(* IEC 61131-3 sources: daoli-st-library/DL_Base (part 17) *)

(* ---- FB_DL_SignalQualify.st ---- *)
(*
  FB_DL_SignalQualify  —  模拟量信号有效性三态联合判定 / Analog signal qualification: over-range, frozen, wire-break
  分类 Category : DL_Base
  版本 Version  : 1.0.0
  来源 Source   : t2-1-lgf-measurement — 信号质量判定族零检索深化
  溯源 Origin   : clean-room 实现，未复制任何源码行
  功能 Function : 1) 对 fRaw 做三态联合判定：超量程（量程域外）/ 断线（低于传感器零点域）/
                  卡死（相邻拍差值持续小于卡死带超过 tFrozenTo），输出 eQual 四态枚举 + bValid；
                  2) 断线判据：fRaw < fScaleLo - fWireMargin（传感器零点域以下）→ eWireBreak；
                  3) 卡死判据：ABS(fRaw - 上拍采样) < fFrozenBand 持续 tFrozenTo → 故障级 03DC；
                  4) bReset 上升沿清全部故障锁存；判定恢复 eOk 沿置信息级码 049E。
  边界 Boundary : ① 组态闸：fScaleLo < fScaleHi 必须成立，违例置故障级 03DB，bValid 强制 FALSE；
                  ② 域判据全部使用当拍量（fRaw 与组态引脚），无锁存量自指；
                  ③ 判定派生链 IF/ELSIF/ELSE 全覆盖，枚举域防御守卫落 03DD 故障锁存；
                  ④ 无 GVL 依赖：纯引脚输入输出，无外部变量引用，无物理 IO 地址。
  依赖 Depends  : 仅 Standard.library（TON / R_TRIG）
  码表 Error codes（段 0001，窗口 03DB~03DD / 049E~04A0）:
    16#0001_03DB 故障级：量程组态非法（fScaleLo >= fScaleHi 或卡死带 <= 0），锁存至 bReset
    16#0001_03DC 故障级：信号卡死超时（冻结判据持续 tFrozenTo），锁存至 bReset
    16#0001_03DD 故障级：判定结果落枚举域外（防御守卫兜底），锁存至 bReset
    16#0001_049E 信息级：信号判定恢复正常（eQual 回 eOk 沿）
    16#0001_049F 信息级：超量程检出（伴随态）
    16#0001_04A0 信息级：断线域命中（伴随态）
  修订历史 Revision :
    2026-11-19  v1.0.0  R41 首版（批次 1 · 序号 1）
*)

TYPE E_DL_SigQual :
(
    eOk        := 0,    // 信号有效，量程域内且动态正常 / Signal valid, in range and dynamic
    eOverRange := 10,   // 超量程：超出组态量程域 / Over range, outside the configured span
    eFrozen    := 20,   // 卡死：变化量持续小于卡死带 / Frozen, change stays below the deadband
    eWireBreak := 30    // 断线：低于传感器零点域 / Wire break, below the sensor zero span
);
END_TYPE

FUNCTION_BLOCK FB_DL_SignalQualify
VAR_INPUT
    fRaw         : LREAL := 0.0;      // 原始采样值 [EU] / Raw sampled value
    fScaleLo     : LREAL := 0.0;      // 量程下限 [EU]，必须 < fScaleHi / Span lower bound
    fScaleHi     : LREAL := 100.0;    // 量程上限 [EU]，必须 > fScaleLo / Span upper bound
    fWireMargin  : LREAL := 1.0;      // 断线判据裕度 [EU]，域 >= 0 / Wire-break margin below span low
    fFrozenBand  : LREAL := 0.01;     // 卡死判定带 [EU]，域 > 0 / Frozen deadband
    tFrozenTo    : TIME := T#5S;      // 卡死确认超时 [ms]，域 > 0 / Frozen confirm timeout
    bReset       : BOOL := FALSE;     // 复位，上升沿清故障锁存 / Reset edge clears fault latches
END_VAR
VAR_OUTPUT
    eQual        : E_DL_SigQual;      // 判定结果出口 / Qualification result
    bValid       : BOOL;              // 判定有效（eOk 且无故障）/ Result usable flag
    bError       : BOOL;              // 故障锁存标志 / Fault latch flag
    nErrId       : UDINT;             // 事件码，0 = 无事件（故障锁存回放优先）/ Event code
END_VAR
VAR
    tonFrozen    : TON;               // 卡死确认定时器，无条件周期刷新 / Frozen confirm timer
    rtReset      : R_TRIG;            // 复位沿实例，无条件周期刷新 / Reset edge instance
    _fLastRaw    : LREAL := 0.0;      // 上拍采样快照 [EU] / Previous scan sample snapshot
    _fDelta      : LREAL;             // 相邻拍差值绝对值 [EU] / Absolute inter-scan delta
    _bFault      : BOOL;              // 故障锁存位（锁存量）/ Latched fault bit
    _uFault      : UDINT;             // 故障码锁存（锁存量）/ Latched fault code
    _uInfo       : UDINT;             // 信息码，每拍重算 / Transient info code
    _bOkPrev     : BOOL;              // 上拍判定有效镜像（恢复沿判据）/ Previous eOk mirror
END_VAR

(* —— 段 0：定时器与沿实例无条件周期刷新（禁置于 IF/CASE 内） —— *)
_fDelta := ABS(fRaw - _fLastRaw);                                       // 相邻拍差值（当拍量）
tonFrozen(IN := (_fDelta < fFrozenBand), PT := tFrozenTo);              // 卡死确认（每拍必调）
rtReset(CLK := bReset);                                                 // 复位沿（每拍必调）

(* —— 段 1：单拍量预清零（锁存量 _bFault/_uFault 不入清单，禁同拍抹除） —— *)
_uInfo := 16#0000_0000;             // 信息码每拍重算
bValid := FALSE;                    // 有效出口缺省 FALSE
nErrId := 16#0000_0000;             // 事件码缺省无事件
eQual := E_DL_SigQual.eOk;          // 判定缺省有效（派生链覆盖改写）

(* —— 段 2：复位沿（唯一故障解除路径，全当拍量） —— *)
IF rtReset.Q THEN                   // rtReset.Q = 当拍量
    _bFault := FALSE;               // 清故障锁存位
    _uFault := 16#0000_0000;        // 清故障锁存码
END_IF

(* —— 段 3：组态域闸（覆盖参与判据换算的全部组态引脚） —— *)
IF (fScaleLo >= fScaleHi) OR (fFrozenBand <= 0.0) OR (TIME_TO_DINT(tFrozenTo) <= 0) THEN
    _uFault := 16#0001_03DB;        // 故障级：量程组态非法
    _bFault := TRUE;
END_IF

(* —— 段 4：三态联合判定（全当拍量判据；派生链 ELSE 兜底 + 枚举域守卫） —— *)
IF NOT _bFault THEN
    IF fRaw < (fScaleLo - ABS(fWireMargin)) THEN
        eQual := E_DL_SigQual.eWireBreak;   // 断线：低于传感器零点域
        _uInfo := 16#0001_04A0;             // 信息级：断线域命中
    ELSIF (fRaw > fScaleHi) OR (fRaw < fScaleLo) THEN
        eQual := E_DL_SigQual.eOverRange;   // 超量程
        _uInfo := 16#0001_049F;             // 信息级：超量程检出
    ELSIF tonFrozen.Q THEN
        eQual := E_DL_SigQual.eFrozen;      // 卡死确认
        _uFault := 16#0001_03DC;            // 故障级：卡死超时
        _bFault := TRUE;
    ELSE
        eQual := E_DL_SigQual.eOk;          // 判定有效
        IF NOT _bOkPrev THEN
            _uInfo := 16#0001_049E;         // 信息级：判定恢复有效沿
        END_IF
    END_IF
    (* 枚举域防御守卫（等价 CASE ELSE 兜底）：判定结果必须落已知枚举域 *)
    IF (eQual <> E_DL_SigQual.eOk) AND (eQual <> E_DL_SigQual.eOverRange)
       AND (eQual <> E_DL_SigQual.eFrozen) AND (eQual <> E_DL_SigQual.eWireBreak) THEN
        _uFault := 16#0001_03DD;            // 故障级：判定态落域外
        _bFault := TRUE;
        eQual := E_DL_SigQual.eOk;          // 强制回已知态
    END_IF
END_IF

(* —— 段 5：出口单点映射（名实同源；故障锁存码回放，禁同拍抹除） —— *)
bValid := (eQual = E_DL_SigQual.eOk) AND (NOT _bFault);   // 有效出口（信息级不置故障）
IF _bFault THEN
    nErrId := _uFault;              // 故障锁存码回放
ELSE
    nErrId := _uInfo;               // 信息码
END_IF
bError := _bFault;                  // 故障标志与锁存位同源
_bOkPrev := (eQual = E_DL_SigQual.eOk);   // 恢复沿判据快照（当拍量快照）
_fLastRaw := fRaw;                  // 上拍采样快照更新（段末统一写）

END_FUNCTION_BLOCK

(* ---- FB_DL_SignalRouteMatrix.st ---- *)
//==============================================================================
// 功能块：FB_DL_SignalRouteMatrix ｜ 中文名称：2×N 可组态信号路由矩阵
// 所属子库：DL_Base ｜ 版本：v1.0.0 ｜ 日期：2026-11-23
// 兼容：CODESYS V3.5+ / TwinCAT 3 / 汇川 InoProShop（纯 IEC 61131-3，零方言）
// 功能描述：2 源 × 4 通道可组态路由矩阵：每通道独立使能 + 来源选择（源 A /
//           源 B / 空置），输出 = 使能 AND 所选源。断源哨兵：存在"通道使能
//           且已选源"但其源信号为 FALSE 时置该源断源哨兵位（正常传递同时
//           留痕，供上层诊断区分"真信号 FALSE"与"通道空置 FALSE"）。
// 开源溯源 (Origin)：原创实现（t2-1-lgf-bitlogic 位逻辑语义深化，零外部源码
//           行，clean-room 独立编写）
// 公开接口清单：输入 aSrcA / aSrcB / {bEnCh1..4, eSelCh1..4}；
//               输出 {bOutCh1..4} / bSrcALost / bSrcBLost / bValid
// 错误码表：无状态机码轨（组合路由无故障级条件）；断源诊断经
//           bSrcALost / bSrcBLost 哨兵位表达，不占用 16#0001 段码位
// 状态机：E_DL_RouteSel（本文件唯一定义，全库唯一属主）：
//           eNone = 0 / eSrcA = 1 / eSrcB = 2；非法选择值走 CASE ELSE 兜底
//           （输出 FALSE 安全侧 + 声明哨兵）
// 边界行为：① 空置通道输出恒 FALSE 且不计入断源哨兵；
//           ② 断源哨兵不屏蔽输出（传递与诊断解耦）；
//           ③ 无定时器/沿实例（纯组合逻辑，无周期刷新义务）；
//           ④ CASE 带 ELSE 非法选择值兜底（输出 FALSE 安全侧）。
// 修订历史：v1.0.0 2026-11-23 首版（R73 派单 · 批 3 · 序 13）
//==============================================================================

(*------------------------------------------------------------------------------
 * 枚举: E_DL_RouteSel（归属本功能块，同文件发布，全库唯一属主）
 * 含义: 通道来源选择，成员与 CASE 标签双向完备。
 *-----------------------------------------------------------------------------*)
TYPE E_DL_RouteSel :
(
    eNone := 0,    // 空置：通道不选源，输出恒 FALSE / Idle, no source selected
    eSrcA := 1,    // 选源 A / Source A selected
    eSrcB := 2     // 选源 B / Source B selected
);
END_TYPE

(*==============================================================================
 * 功能块: FB_DL_SignalRouteMatrix
 * 调用约定: 每个扫描周期无条件调用一次；纯组合路由，无跨拍驻留状态。
 *==============================================================================*)
FUNCTION_BLOCK FB_DL_SignalRouteMatrix
VAR_INPUT
    aSrcA   : BOOL := FALSE;           // 源 A 信号 [—] / Source A signal
    aSrcB   : BOOL := FALSE;           // 源 B 信号 [—] / Source B signal
    bEnCh1  : BOOL := FALSE;           // 通道 1 使能 / Channel 1 enable
    eSelCh1 : E_DL_RouteSel := E_DL_RouteSel.eNone; // 通道 1 来源选择 / Channel 1 source select
    bEnCh2  : BOOL := FALSE;           // 通道 2 使能 / Channel 2 enable
    eSelCh2 : E_DL_RouteSel := E_DL_RouteSel.eNone; // 通道 2 来源选择 / Channel 2 source select
    bEnCh3  : BOOL := FALSE;           // 通道 3 使能 / Channel 3 enable
    eSelCh3 : E_DL_RouteSel := E_DL_RouteSel.eNone; // 通道 3 来源选择 / Channel 3 source select
    bEnCh4  : BOOL := FALSE;           // 通道 4 使能 / Channel 4 enable
    eSelCh4 : E_DL_RouteSel := E_DL_RouteSel.eNone; // 通道 4 来源选择 / Channel 4 source select
END_VAR
VAR_OUTPUT
    bOutCh1 : BOOL;                    // 通道 1 路由输出 / Channel 1 routed output
    bOutCh2 : BOOL;                    // 通道 2 路由输出 / Channel 2 routed output
    bOutCh3 : BOOL;                    // 通道 3 路由输出 / Channel 3 routed output
    bOutCh4 : BOOL;                    // 通道 4 路由输出 / Channel 4 routed output
    bSrcALost : BOOL;                  // 断源哨兵：有通道选 A 但源 A 为 FALSE / Source-A lost sentinel
    bSrcBLost : BOOL;                  // 断源哨兵：有通道选 B 但源 B 为 FALSE / Source-B lost sentinel
    bValid  : BOOL;                    // 输出可用标志 / Outputs usable flag
END_VAR

// ---- 段 0｜出口默认值：哨兵每拍重算（组合诊断位不锁存）----
bSrcALost := FALSE;                   // 源 A 断源哨兵先清零 / Source-A lost sentinel cleared first
bSrcBLost := FALSE;                   // 源 B 断源哨兵先清零 / Source-B lost sentinel cleared first
bValid    := TRUE;                    // 可用标志默认 TRUE / Usable flag preset TRUE

// ---- 段 1｜通道 1/2 路由（CASE 带 ELSE；空置与非法值安全侧输出 FALSE）----
CASE eSelCh1 OF                       // 通道 1 来源判决 / Channel 1 source decision
    E_DL_RouteSel.eNone:               // 空置：输出 FALSE，不计哨兵 / Idle, FALSE, no sentinel
        bOutCh1 := FALSE;              // 通道 1 输出 / Channel 1 output
    E_DL_RouteSel.eSrcA:               // 选源 A：使能闸 + 断源哨兵留痕 / Source A, enable gate plus lost sentinel
        bOutCh1 := bEnCh1 AND aSrcA;   // 通道 1 输出 / Channel 1 output
        bSrcALost := bSrcALost OR (bEnCh1 AND NOT aSrcA); // 断源哨兵累积 / Lost sentinel accumulate
    E_DL_RouteSel.eSrcB:               // 选源 B：使能闸 + 断源哨兵留痕 / Source B, enable gate plus lost sentinel
        bOutCh1 := bEnCh1 AND aSrcB;   // 通道 1 输出 / Channel 1 output
        bSrcBLost := bSrcBLost OR (bEnCh1 AND NOT aSrcB); // 断源哨兵累积 / Lost sentinel accumulate
    ELSE                               // 非法选择值兜底（R21：CASE 必带 ELSE）
        bOutCh1 := FALSE;              // 安全侧输出 FALSE / Safe-side FALSE output
END_CASE
CASE eSelCh2 OF                       // 通道 2 来源判决 / Channel 2 source decision
    E_DL_RouteSel.eNone:               // 空置：输出 FALSE，不计哨兵 / Idle, FALSE, no sentinel
        bOutCh2 := FALSE;              // 通道 2 输出 / Channel 2 output
    E_DL_RouteSel.eSrcA:               // 选源 A：使能闸 + 断源哨兵留痕 / Source A, enable gate plus lost sentinel
        bOutCh2 := bEnCh2 AND aSrcA;   // 通道 2 输出 / Channel 2 output
        bSrcALost := bSrcALost OR (bEnCh2 AND NOT aSrcA); // 断源哨兵累积 / Lost sentinel accumulate
    E_DL_RouteSel.eSrcB:               // 选源 B：使能闸 + 断源哨兵留痕 / Source B, enable gate plus lost sentinel
        bOutCh2 := bEnCh2 AND aSrcB;   // 通道 2 输出 / Channel 2 output
        bSrcBLost := bSrcBLost OR (bEnCh2 AND NOT aSrcB); // 断源哨兵累积 / Lost sentinel accumulate
    ELSE                               // 非法选择值兜底（R21：CASE 必带 ELSE）
        bOutCh2 := FALSE;              // 安全侧输出 FALSE / Safe-side FALSE output
END_CASE

// ---- 段 2｜通道 3/4 路由（同段 1 口径）----
CASE eSelCh3 OF                       // 通道 3 来源判决 / Channel 3 source decision
    E_DL_RouteSel.eNone:               // 空置：输出 FALSE，不计哨兵 / Idle, FALSE, no sentinel
        bOutCh3 := FALSE;              // 通道 3 输出 / Channel 3 output
    E_DL_RouteSel.eSrcA:               // 选源 A：使能闸 + 断源哨兵留痕 / Source A, enable gate plus lost sentinel
        bOutCh3 := bEnCh3 AND aSrcA;   // 通道 3 输出 / Channel 3 output
        bSrcALost := bSrcALost OR (bEnCh3 AND NOT aSrcA); // 断源哨兵累积 / Lost sentinel accumulate
    E_DL_RouteSel.eSrcB:               // 选源 B：使能闸 + 断源哨兵留痕 / Source B, enable gate plus lost sentinel
        bOutCh3 := bEnCh3 AND aSrcB;   // 通道 3 输出 / Channel 3 output
        bSrcBLost := bSrcBLost OR (bEnCh3 AND NOT aSrcB); // 断源哨兵累积 / Lost sentinel accumulate
    ELSE                               // 非法选择值兜底（R21：CASE 必带 ELSE）
        bOutCh3 := FALSE;              // 安全侧输出 FALSE / Safe-side FALSE output
END_CASE
CASE eSelCh4 OF                       // 通道 4 来源判决 / Channel 4 source decision
    E_DL_RouteSel.eNone:               // 空置：输出 FALSE，不计哨兵 / Idle, FALSE, no sentinel
        bOutCh4 := FALSE;              // 通道 4 输出 / Channel 4 output
    E_DL_RouteSel.eSrcA:               // 选源 A：使能闸 + 断源哨兵留痕 / Source A, enable gate plus lost sentinel
        bOutCh4 := bEnCh4 AND aSrcA;   // 通道 4 输出 / Channel 4 output
        bSrcALost := bSrcALost OR (bEnCh4 AND NOT aSrcA); // 断源哨兵累积 / Lost sentinel accumulate
    E_DL_RouteSel.eSrcB:               // 选源 B：使能闸 + 断源哨兵留痕 / Source B, enable gate plus lost sentinel
        bOutCh4 := bEnCh4 AND aSrcB;   // 通道 4 输出 / Channel 4 output
        bSrcBLost := bSrcBLost OR (bEnCh4 AND NOT aSrcB); // 断源哨兵累积 / Lost sentinel accumulate
    ELSE                               // 非法选择值兜底（R21：CASE 必带 ELSE）
        bOutCh4 := FALSE;              // 安全侧输出 FALSE / Safe-side FALSE output
END_CASE

// ---- 段 3｜统一出口：可用标志（纯组合无防御失败路径）----
bValid := TRUE;                       // 组合路由恒可用 / Combinational routing always usable
END_FUNCTION_BLOCK

(* ---- FB_DL_SignalSeqGuard.st ---- *)
(*
  ==================================================================
  组件名 Component  : FB_DL_SignalSeqGuard
  分类   Category   : DL_Base
  复杂度 Complexity  : cx3
  版本   Version    : 1.0.0
  功能   Purpose    : 多路信号到达顺序守卫。N = 4 路布尔信号按期望序（ENUM 四选一：
                      升序 1→2→3→4 / 降序 4→3→2→1 / 对 1→2 / 对 3→4）在 tWindow
                      内逐沿校验到达顺序；乱序即置 eFault = eOrderViolation 并锁存，
                      窗内未完成置 eWindowTimeout；正常序完成置 bSeqOk 单拍脉冲。
                      复位上升沿清全部锁存。同拍多沿按 1..4 固定序检查（确定性口径）。
  来源   Source     : t2-1-lgf-converter
  溯源   Origin     : IEC 61131-3 标准语义的道莅防御性实现；到达顺序校验为通用
                      联锁语义，clean-room 自研实现，未复制任何闭源代码行。
  平台   Platform   : 纯 IEC 61131-3（TON / R_TRIG / ARRAY，无私有库）
  作者   Author     : 道莅代码库 · PLC 编程专家（R56）
  ------------------------------------------------------------------
  边界 Boundary     :
                      一 本件只做到达顺序校验，不产生任何输出命令（属主边界）；
                      二 eWait 类相（eRun）退出条件 ≥2 条：完成沿 / 超时 / 乱序 /
                         失能，四条并列（R98）；
                      三 序列表在组态相一次性落定，乱序判据只用序表与步进游标；
                      四 故障锁存解除路径 = bReset 上升沿（唯一路径，头注释声明，R188）；
                      五 无全局变量、无外部变量声明、无物理地址寻址。
  输出契约 Output contract:
                      bSeqOk 为单拍脉冲（内部 _bOkInt 置位、统一出口映射后撤销，R187）；
                      eFault 为锁存回放；eModeBad 为模式枚举非法兜底（R128）。
  修订记录 Revision  :
    2026-11-20  v1.0.0  R56 首版（批 2 · 序号 7）
  ==================================================================
*)

TYPE E_DL_SsgMode :
(
    eAscending  := 0, // 升序：1→2→3→4 / ascending, one to four
    eDescending := 1, // 降序：4→3→2→1 / descending, four to one
    ePair12     := 2, // 对序：1→2 / pair order, one then two
    ePair34     := 3  // 对序：3→4 / pair order, three then four
);
END_TYPE

TYPE E_DL_SsgPhase :
(
    eIdle  := 0,  // 空闲：等待启动 / idle, waiting for the start
    eRun   := 10, // 校验中：逐沿核对到达顺序 / running, the arrivals are checked edge by edge
    eDone  := 20, // 完成：顺序通过，驻留一拍 / done, the order passed and the phase holds one scan
    eFault := 90  // 故障：成因锁存 / fault, the cause is latched
);
END_TYPE

TYPE E_DL_SsgFault :
(
    eNone          := 0, // 无成因 / no cause
    eOrderViolation:= 1, // 到达顺序违例（故障级，与 bError 配对）/ the arrival order was violated, fault grade paired with bError
    eWindowTimeout := 2, // 时窗内未完成（故障级，与 bError 配对）/ the window expired without completion, fault grade paired with bError
    eModeBad       := 3, // 模式枚举非法（故障级，与 bError 配对）/ the mode enumeration is illegal, fault grade paired with bError
    ePhaseBad      := 4  // 非法相位兜底（故障级，与 bError 配对）/ illegal phase fallback, fault grade paired with bError
);
END_TYPE

FUNCTION_BLOCK FB_DL_SignalSeqGuard
VAR_INPUT
    bEnable   : BOOL := TRUE;    // 使能，失能时停校验回空闲 [-] / enable, the check stops when disabled
    bReset    : BOOL := FALSE;   // 复位上升沿清全部锁存 [-] / reset rising edge clears every latch
    bIn1      : BOOL := FALSE;   // 信号 1 [-] / signal one
    bIn2      : BOOL := FALSE;   // 信号 2 [-] / signal two
    bIn3      : BOOL := FALSE;   // 信号 3 [-] / signal three
    bIn4      : BOOL := FALSE;   // 信号 4 [-] / signal four
    eSeqMode  : E_DL_SsgMode := E_DL_SsgMode.eAscending; // 期望到达序 [枚举] / the expected arrival order [enum]
    tWindow   : TIME := T#2S;    // 到达顺序时窗 [毫秒]，域 大于零 / arrival order window [millisecond], domain above zero
END_VAR
VAR_OUTPUT
    bSeqOk    : BOOL := FALSE; // 顺序通过单拍脉冲 [-] / the order passed single shot pulse
    nStep     : INT := 0;      // 已到位步数 [步] / the arrived step count [step]
    ePhase    : E_DL_SsgPhase := E_DL_SsgPhase.eIdle; // 相位出口 [枚举] / phase outlet [enum]
    eFault    : E_DL_SsgFault := E_DL_SsgFault.eNone; // 成因出口，锁存回放 [枚举] / cause outlet replayed from the latch [enum]
    bError    : BOOL := FALSE; // 故障锁存标志 [-] / fault latch flag
END_VAR
VAR
    rtIn1     : R_TRIG;  // 信号 1 沿检测，段 0 无条件刷新 / signal one edge, refreshed unconditionally in segment zero
    rtIn2     : R_TRIG;  // 信号 2 沿检测，段 0 无条件刷新 / signal two edge, refreshed unconditionally in segment zero
    rtIn3     : R_TRIG;  // 信号 3 沿检测，段 0 无条件刷新 / signal three edge, refreshed unconditionally in segment zero
    rtIn4     : R_TRIG;  // 信号 4 沿检测，段 0 无条件刷新 / signal four edge, refreshed unconditionally in segment zero
    rtReset   : R_TRIG;  // 复位沿检测，段 0 无条件刷新 / reset edge, refreshed unconditionally in segment zero
    tonWindow : TON;     // 到达顺序时窗，段 0 无条件刷新 / arrival window timer, refreshed unconditionally in segment zero
    _ePhase   : E_DL_SsgPhase := E_DL_SsgPhase.eIdle; // 内部相位，CASE 唯一写入目标 / internal phase, the only CASE write target
    _eFaulC   : E_DL_SsgFault := E_DL_SsgFault.eNone; // 故障级成因，锁存至复位沿 / fault cause, latched until the reset edge
    _bFault   : BOOL := FALSE; // 故障锁存位 [-] / fault latch bit
    _bInit    : BOOL := FALSE; // 首扫初始化完成标志（R310）/ first scan initialisation flag
    _bOkInt   : BOOL := FALSE; // 通过脉冲内部位，统一出口映射 / internal passed bit, mapped at the unified outlet
    _nStep    : INT := 0;      // 已到位步数 [步] / the arrived step count [step]
    _nSeqLen  : INT := 4;      // 序列长度（四序或两序）[步] / the sequence length, four or two steps
    _nSig     : INT := 0;      // 本拍到沿的信号号 [信号号] / the signal number that edged this scan
    _anOrder  : ARRAY[1..4] OF INT := [0, 0, 0, 0]; // 期望到达序表（0 = 空槽）[信号号] / the expected order table, zero is an empty slot
END_VAR

// 段 0｜定时器与沿检测无条件周期刷新（禁入分支），IN 只串相位闸与故障闸（FB50-1）/ segment 0, unconditional refresh, no instance call inside a branch
rtIn1(CLK := bIn1); // 信号 1 沿 / the signal one edge
rtIn2(CLK := bIn2); // 信号 2 沿 / the signal two edge
rtIn3(CLK := bIn3); // 信号 3 沿 / the signal three edge
rtIn4(CLK := bIn4); // 信号 4 沿 / the signal four edge
rtReset(CLK := bReset); // 复位沿 / the reset edge
tonWindow(IN := (_ePhase = E_DL_SsgPhase.eRun) AND (NOT _bFault), PT := tWindow); // 到达顺序时窗，IN 串校验相闸与故障闸 / the arrival window with the phase and fault gates on IN

// 段 1｜首扫初始化（R310）/ segment 1, first scan initialisation
IF NOT _bInit THEN // 首扫一拍 / the very first scan
    _bInit := TRUE; // 置首扫完成标志 / raise the first scan flag
    _ePhase := E_DL_SsgPhase.eIdle; // 相位从空闲起步 / the phase starts from idle
    _eFaulC := E_DL_SsgFault.eNone; // 故障级成因清零 / clear the fault cause
    _bFault := FALSE; // 故障锁存清零 / clear the fault latch
    _nStep := 0; // 步数清零 / clear the step count
END_IF

// 段 2｜复位沿作用域：清锁存 / 迁相位 / 清步数（三项逐项声明）/ segment 2, reset edge scope declared item by item
IF rtReset.Q THEN // 复位沿 / the reset edge
    _bFault := FALSE; // 作用域一：清故障锁存 / scope one, clear the fault latch
    _eFaulC := E_DL_SsgFault.eNone; // 作用域一：清故障级成因 / scope one, clear the fault cause
    _ePhase := E_DL_SsgPhase.eIdle; // 作用域二：迁回空闲相 / scope two, migrate back to idle
    _nStep := 0; // 作用域三：清步数 / scope three, clear the step count
END_IF

// 段 3｜序表组态：按模式一次性落定，非法模式判故障 / segment 3, the order table settles per the mode, an illegal mode faults
CASE eSeqMode OF // 模式分派 / the mode dispatch
E_DL_SsgMode.eAscending: // 升序 / ascending
    _anOrder[1] := 1; // 第一位信号 1 / the first slot takes signal one
    _anOrder[2] := 2; // 第二位信号 2 / the second slot takes signal two
    _anOrder[3] := 3; // 第三位信号 3 / the third slot takes signal three
    _anOrder[4] := 4; // 第四位信号 4 / the fourth slot takes signal four
    _nSeqLen := 4; // 序列长度四 / the length is four
E_DL_SsgMode.eDescending: // 降序 / descending
    _anOrder[1] := 4; // 第一位信号 4 / the first slot takes signal four
    _anOrder[2] := 3; // 第二位信号 3 / the second slot takes signal three
    _anOrder[3] := 2; // 第三位信号 2 / the third slot takes signal two
    _anOrder[4] := 1; // 第四位信号 1 / the fourth slot takes signal one
    _nSeqLen := 4; // 序列长度四 / the length is four
E_DL_SsgMode.ePair12: // 对序 1→2 / pair one then two
    _anOrder[1] := 1; // 第一位信号 1 / the first slot takes signal one
    _anOrder[2] := 2; // 第二位信号 2 / the second slot takes signal two
    _anOrder[3] := 0; // 空槽 / an empty slot
    _anOrder[4] := 0; // 空槽 / an empty slot
    _nSeqLen := 2; // 序列长度二 / the length is two
E_DL_SsgMode.ePair34: // 对序 3→4 / pair three then four
    _anOrder[1] := 3; // 第一位信号 3 / the first slot takes signal three
    _anOrder[2] := 4; // 第二位信号 4 / the second slot takes signal four
    _anOrder[3] := 0; // 空槽 / an empty slot
    _anOrder[4] := 0; // 空槽 / an empty slot
    _nSeqLen := 2; // 序列长度二 / the length is two
ELSE // 非法模式兜底（R128）/ the illegal mode fallback
    IF (NOT _bFault) AND (_ePhase <> E_DL_SsgPhase.eFault) THEN // 未锁存才迁移（防同拍抹除）/ migrate only while unlatched
        _bFault := TRUE; // 置故障锁存 / raise the fault latch
        _eFaulC := E_DL_SsgFault.eModeBad; // 故障级成因（R45 配对 bError）/ the fault cause paired with bError
        _ePhase := E_DL_SsgPhase.eFault; // 迁故障相 / migrate to the fault phase
    END_IF
END_CASE

// 段 4｜本拍到沿信号号判定：同拍多沿按 1..4 固定序（确定性口径）/ segment 4, the edged signal number, multiple edges resolve in the fixed one to four order
_nSig := 0; // 信号号预置零 / preset the signal number to zero
IF rtIn1.Q THEN // 信号 1 到沿 / signal one edged
    _nSig := 1; // 记信号 1 / take signal one
ELSIF rtIn2.Q THEN // 信号 2 到沿 / signal two edged
    _nSig := 2; // 记信号 2 / take signal two
ELSIF rtIn3.Q THEN // 信号 3 到沿 / signal three edged
    _nSig := 3; // 记信号 3 / take signal three
ELSIF rtIn4.Q THEN // 信号 4 到沿 / signal four edged
    _nSig := 4; // 记信号 4 / take signal four
END_IF

// 段 5｜相位机：ENUM + CASE，含 ELSE 非法相位兜底（R128）/ segment 5, the phase machine with an ELSE fallback
CASE _ePhase OF
E_DL_SsgPhase.eIdle: // 空闲相：使能且无故障即起校验 / idle, the check starts when enabled and unfaulted
    IF bEnable AND (NOT _bFault) THEN // 使能且无故障 / enabled and unfaulted
        _nStep := 0; // 步数清零 / clear the step count
        _ePhase := E_DL_SsgPhase.eRun; // 迁校验相 / migrate to the run phase
    END_IF

E_DL_SsgPhase.eRun: // 校验相：逐沿核对到达顺序（退出条件 ≥2：完成 / 超时 / 乱序 / 失能，R98）/ the run phase with at least two exit conditions
    nStep := _nStep; // 步数出口跟随 / the step outlet follows
    IF NOT bEnable THEN // 失能 / disabled
        _ePhase := E_DL_SsgPhase.eIdle; // 回空闲相 / return to idle
    ELSIF tonWindow.Q THEN // 时窗耗尽未完成 / the window expired without completion
        _bFault := TRUE; // 置故障锁存 / raise the fault latch
        _eFaulC := E_DL_SsgFault.eWindowTimeout; // 故障级成因（R45 配对 bError）/ the fault cause paired with bError
        _ePhase := E_DL_SsgPhase.eFault; // 迁故障相 / migrate to the fault phase
    ELSIF _nSig > 0 THEN // 本拍有信号到沿 / a signal edged this scan
        IF _nSig = _anOrder[_nStep + 1] THEN // 与期望序位一致 / the arrival matches the expected slot
            _nStep := _nStep + 1; // 步数推进 / advance the step
            IF _nStep >= _nSeqLen THEN // 序列完成 / the sequence is complete
                _bOkInt := TRUE; // 通过脉冲内部位置位（统一出口映射，R187）/ raise the internal passed bit, mapped at the unified outlet
                _ePhase := E_DL_SsgPhase.eDone; // 迁完成相 / migrate to the done phase
            END_IF
        ELSE // 乱序 / an out of order arrival
            _bFault := TRUE; // 置故障锁存 / raise the fault latch
            _eFaulC := E_DL_SsgFault.eOrderViolation; // 故障级成因（R45 配对 bError）/ the fault cause paired with bError
            _ePhase := E_DL_SsgPhase.eFault; // 迁故障相 / migrate to the fault phase
        END_IF
    END_IF

E_DL_SsgPhase.eDone: // 完成相：脉冲已交付（拍 N 进入：序到位 / 本拍行为：脉冲映射 / 拍 N+1 转出：无条件回空闲，R80 三段）/ the done phase, the pulse was delivered
    _ePhase := E_DL_SsgPhase.eIdle; // 无条件回空闲相准备下一轮（失能态下同样回到空闲语义）/ back to idle for the next round unconditionally, the same idle semantics under a disable

E_DL_SsgPhase.eFault: // 故障相：成因锁存，等待复位沿 / the fault phase, the cause is latched until the reset edge
    nStep := _nStep; // 步数出口冻结保持 / the step outlet holds frozen

ELSE // 非法相位兜底（R128）/ the illegal phase fallback
    _bFault := TRUE; // 置故障锁存 / raise the fault latch
    _eFaulC := E_DL_SsgFault.ePhaseBad; // 故障级成因（R45 配对 bError）/ the fault cause paired with bError
    _ePhase := E_DL_SsgPhase.eFault; // 迁故障相 / migrate to the fault phase
END_CASE

// 段 6｜统一出口 / segment 6, the unified outlet
bSeqOk := _bOkInt; // 通过脉冲映射本拍值 / map the passed pulse for this scan
_bOkInt := FALSE; // 映射后立即撤销，保证单拍宽度（R187 两段式）/ revoke right after mapping to keep a single scan width
nStep := _nStep; // 步数出口 / the step outlet
ePhase := _ePhase; // 相位出口单点映射 / single point phase outlet mapping
eFault := _eFaulC; // 成因出口锁存回放 / the cause outlet replayed from the latch
bError := _bFault; // 故障标志与锁存位同源 / the fault flag shares the latch source
END_FUNCTION_BLOCK

(* ---- FB_DL_SignalStagnationWatch.st ---- *)
(*
  ==================================================================
  组件名 Component  : FB_DL_SignalStagnationWatch
  分类   Category   : DL_Base
  复杂度 Complexity  : cx3
  版本   Version    : 1.0.0
  功能   Purpose    : 信号呆滞（卡死）检测。双判据持续 tStall 判呆滞：
                      ① 值纹波消失——相邻拍变化量 |Δ| ≤ fEps 持续；
                      ② 伴生活动信号边沿计数归零——活动观测窗内零边沿。
                      两判据同时成立才出呆滞电平与单拍事件。
  来源   Source     : iec-std-wrapper（T0）
  溯源   Origin     : IEC 61131-3 标准语义的道莅防御性实现；呆滞双判据为公开
                      诊断语义，clean-room 自研实现，未复制任何闭源代码行。
  平台   Platform   : 纯 IEC 61131-3（Standard.library: TON / R_TRIG，无私有库）
  分工声明 Split     : 与 FB_DL_SignalDebounce 分工——Debounce 是（抑制）件
                      （吸收毛刺防误动），本件是（检出）件（发现信号呆滞
                      疑点），方向相反、互不替代；与 FB_DL_SensorDropoutHold
                      分工——掉线保持件处理无效值，本件处理有效但不动值。
  作者   Author     : 道莅代码库 · PLC 编程专家（R57）
  ------------------------------------------------------------------
  边界 Boundary     :
                      一 fEps 为显式纹波死区参数，组态闸要求 > 0（信息级）；
                      二 tStall 期间边沿计数窗独立自复位（R188：IN := NOT Q），
                         与呆滞计时互不牵连；
                      三 使能断开即复位：计时清零、窗计数清零、出口回假，
                         不锁存（每拍重算）；
                      四 首扫快照取当拍，无假呆滞（tonStall 从零起步）；
                      五 无全局变量、无外部变量声明、无物理地址寻址。
  修订记录 Revision  :
    2026-11-21  v1.0.0  R57 首版（批 1 · 序号 4）
  ==================================================================
*)

FUNCTION_BLOCK FB_DL_SignalStagnationWatch
VAR_INPUT
    fValue    : LREAL := 0.0;    // 被监视值 [工程单位] / the monitored value [engineering unit]
    bActivity : BOOL := FALSE;   // 伴生活动信号（如传感器自检翻转）[-] / the companion activity signal
    fEps      : LREAL := 0.01;   // 纹波死区 [工程单位]，域 大于零 / the ripple deadband [engineering unit], above zero
    tStall    : TIME := T#10S;   // 呆滞确认窗 [毫秒] / the stall confirm window [millisecond]
    tEdgeWin  : TIME := T#5S;    // 边沿观测窗 [毫秒] / the edge observation window [millisecond]
    bEnable   : BOOL := TRUE;    // 使能，失能即复位不锁存 [-] / enable, disabling resets without latching
    bReset    : BOOL := FALSE;   // 复位上升沿清计数 [-] / reset rising edge clears the counters
END_VAR
VAR_OUTPUT
    bStalled    : BOOL := FALSE; // 呆滞电平出口（双判据同时成立）[-] / the stalled level outlet, both criteria met
    bStallEvent : BOOL := FALSE; // 呆滞进入单拍事件 [-] / the stall entry one-scan event
    nRippleCnt  : UDINT := 0;    // 纹波事件累计 [次] / the ripple event count [count]
    nActWinCnt  : UDINT := 0;    // 当前观测窗内活动边沿计数 [次] / the activity edge count in the current window [count]
    uErrorId    : UDINT := 0;    // 信息级码，0 = 正常 / informational code, zero is ok
    bError      : BOOL := FALSE; // 信息级错误标志（每拍重算）/ informational flag, recomputed each scan
END_VAR
VAR
    rtReset : R_TRIG;  // 复位沿检测，段 0 无条件刷新 / the reset edge, refreshed unconditionally
    rtAct   : R_TRIG;  // 活动信号沿检测，段 0 无条件刷新 / the activity edge, refreshed unconditionally
    rtStall : R_TRIG;  // 呆滞电平沿检测，段 0 无条件刷新 / the stalled level edge, refreshed unconditionally
    tonStall: TON;     // 呆滞确认窗，段 0 无条件刷新 / the stall confirm timer, refreshed unconditionally
    tonWin  : TON;     // 边沿观测窗（自复位），段 0 无条件刷新 / the observation window, self resetting, refreshed unconditionally
    _bInit  : BOOL := FALSE; // 首扫初始化完成标志（R310）/ first scan flag
    _fPrev  : LREAL := 0.0;  // 上拍值快照 [工程单位] / previous scan value snapshot [engineering unit]
    _bRipple: BOOL := FALSE; // 本拍纹波事件标记（上拍值供段 0 判据闸使用）/ the ripple flag this scan, the last value feeds the segment zero gate
    _bCfgOk : BOOL := FALSE; // 组态域内 [-] / the configuration inside the domain
END_VAR

// 段 0｜定时器与沿检测无条件周期刷新（禁入分支）；观测窗自复位（R188）/ segment 0, unconditional refresh, the window self resetting
rtReset(CLK := bReset); // 复位沿 / the reset edge
rtAct(CLK := bActivity); // 活动沿 / the activity edge
rtStall(CLK := bStalled); // 呆滞电平沿 / the stalled level edge
tonStall(IN := _bCfgOk AND bEnable AND (NOT _bRipple) AND (rtAct.Q = FALSE) AND (nActWinCnt = 0), PT := tStall); // 呆滞窗，IN 串双判据闸 / the stall timer gated by both criteria
tonWin(IN := bEnable AND (NOT tonWin.Q), PT := tEdgeWin); // 观测窗自复位循环（R188）/ the self resetting observation loop

// 段 1｜首扫初始化（R310）：快照取当拍防假呆滞 / segment 1, first scan, the snapshot takes this scan
IF NOT _bInit THEN // 首扫一拍 / the first scan
    _bInit := TRUE; // 置首扫标志 / raise the flag
    _fPrev := fValue; // 快照取当拍 / the snapshot takes this scan
END_IF

// 段 2｜复位沿作用域：清计数（出口电平随计时自清，无需另清）/ segment 2, reset edge scope
IF rtReset.Q THEN // 复位沿 / the reset edge
    nRippleCnt := 0; // 清纹波计数 / clear the ripple counter
    nActWinCnt := 0; // 清窗计数 / clear the window counter
END_IF

// 段 3｜组态域闸（信息级，每拍重算）/ segment 3, the configuration gate, informational
_bCfgOk := (fEps > 0.0) AND (fEps = fEps) AND ((fEps - fEps) = (fEps - fEps)) AND (tStall > T#0S) AND (tEdgeWin > T#0S); // 死区与窗域判定 / the deadband and window verdict
IF NOT _bCfgOk THEN // 组态非法 / an illegal configuration
    uErrorId := 16#0001_0001; // 信息级：组态越域 / informational, a config violation
    bError   := TRUE; // 置信息级标志 / raise the flag
ELSE // 域内 / inside the domain
    uErrorId := 16#0000_0000; // 正常码 / the ok code
    bError   := FALSE; // 清标志 / clear the flag
END_IF

// 段 4｜双判据量测 / segment 4, the dual criteria measurement
_bRipple := ABS(fValue - _fPrev) > fEps; // 纹波判据（变化量超死区）/ the ripple verdict beyond the deadband
IF _bRipple THEN // 纹波事件 / a ripple event
    nRippleCnt := nRippleCnt + 1; // 纹波计数推进 / advance the ripple counter
    IF nRippleCnt = 4294967295 THEN // UDINT 上界防回绕 / the wrap guard
        nRippleCnt := 4294967294; // 钳在次上界 / clamp below the ceiling
    END_IF
END_IF
IF rtAct.Q THEN // 活动沿 / an activity edge
    nActWinCnt := nActWinCnt + 1; // 窗内计数推进 / advance the window counter
END_IF
IF tonWin.Q THEN // 观测窗到期：窗计数独立归零重开（边界二）/ the window expired, the counter reset independently
    nActWinCnt := 0; // 窗计数归零 / the window counter zeroed
END_IF
IF NOT bEnable THEN // 失能即复位不锁存（边界三）/ disabled resets without latching
    nRippleCnt := 0; // 清纹波计数 / clear the ripple counter
    nActWinCnt := 0; // 清窗计数 / clear the window counter
END_IF

// 段 5｜统一出口：双判据电平 + 进入事件 / segment 5, the unified outlet
bStalled := _bCfgOk AND bEnable AND tonStall.Q AND (nActWinCnt = 0); // 双判据电平 / the dual criteria level
bStallEvent := rtStall.Q; // 进入单拍事件（沿检测已无条件刷新）/ the entry one-scan event
IF NOT bEnable THEN // 失能拍出口回假 / the disabled scan forces false
    bStalled := FALSE; // 电平回假 / the level false
    bStallEvent := FALSE; // 事件回假 / the event false
END_IF
_fPrev := fValue; // 快照推进（无条件）/ the snapshot advances unconditionally
END_FUNCTION_BLOCK

(* ---- FB_DL_SignalStuckWatch.st ---- *)
(*
  Name        : FB_DL_SignalStuckWatch
  Category    : DL_Base
  Version     : 1.0.0
  Purpose     : 信号卡死监视：监视值在卡死判定窗内变化量始终不超过死区（变化率恒零）即报警，捕捉传感器冻结/线束搭死；/ Signal stuck watch: raises an alarm when the monitored value stays within the deadband for the whole stuck window, catching frozen sensors or shorted wiring
  溯源        : 借 t2-1-lgf 的分类/参数域组织，clean-room 实现
  Boundary    : ① 组态闸：死区 < 0 / 卡死窗 <= T#0S → 锁存故障（死区 0 合法：严格等值判死）；
                ② 卡死判定窗用 TON，IN 由「未变化 + 已取基线」派生并串 eMon 相位闸（族③：eIdle/eFault 不计时，上拍相位 1 拍延迟可接受），段 0 无 IF 包裹；
                ③ 非有限值该拍不更新基线不计时（防 NaN 把窗持续清零而漏报，也防污染基线）；
                ④ 基线快照在迁入 eMon 拍取（fValue 首值），变化超死区即刷新基线并重置计时；
                ⑤ bStuck 锁存至复位沿；bStuck 起始沿单拍脉冲 bStuckEdge 供事件记录（R187 两段式）。
*)
TYPE E_DL_SswState :
(
    eIdle  := 0,                             (* 未使能 / Disabled *)
    eMon   := 10,                            (* 卡死监视运行 / Monitoring *)
    eFault := 90                             (* 故障锁存相 / Fault latched *)
);
END_TYPE

TYPE E_DL_SswCause :
(
    eNone       := 0,                        (* 无故障成因 / No cause *)
    eCfgIllegal := 1,                        (* 组态非法：死区/窗口越域 / Illegal config *)
    eStuck      := 2,                        (* 信号卡死（窗满无有效变化） / Signal stuck *)
    ePhaseBad   := 3                         (* 非法相位兜底 / Illegal phase fallback *)
);
END_TYPE

FUNCTION_BLOCK FB_DL_SignalStuckWatch
VAR_INPUT
    fValue    : REAL := 0.0;                 (* 被监视信号值（任意工程量）[-] / Monitored signal value *)
    fDeadband : REAL := 0.01;               (* 变化判定死区，域 >= 0 [工程单位] / Deadband for change detection *)
    tStuckWin : TIME := T#60S;              (* 卡死判定窗长，域 > T#0S [ms] / Stuck window length, > 0 *)
    bEnable   : BOOL := TRUE;               (* 监视使能 [-] / Enable *)
    bReset    : BOOL := FALSE;              (* 复位命令，上升沿清报警与故障 [-] / Reset command *)
END_VAR
VAR_OUTPUT
    fDelta    : REAL;                        (* 本拍相对基线变化量（实时派生）[工程单位] / Delta versus baseline *)
    bStuck    : BOOL;                        (* 卡死报警锁存（复位沿清）[-] / Stuck alarm latched *)
    bStuckEdge: BOOL;                        (* 卡死报警起始沿（单拍脉冲）[-] / Stuck alarm rising edge pulse *)
    fLastMove : TIME;                       (* 最近一次有效变化距今时长（本窗计时镜像）[ms] / Time since last valid move *)
    eState    : E_DL_SswState;               (* 状态出口 / State outlet *)
    eCause    : E_DL_SswCause;               (* 故障成因出口（R190 归因唯一） / Fault cause outlet *)
    bError    : BOOL;                        (* 故障锁存标志 [-] / Fault latch flag *)
END_VAR
VAR
    _eState   : E_DL_SswState := E_DL_SswState.eIdle;    (* 内部相位（CASE 唯一写入目标） / Internal phase *)
    _eCause   : E_DL_SswCause := E_DL_SswCause.eNone;    (* 故障成因锁存量 / Latched cause *)
    rtReset   : R_TRIG;                      (* 复位沿实例，段 0 无条件调用 / Reset edge instance *)
    rtStuck   : R_TRIG;                      (* 卡死计时器输出沿实例，段 0 无条件调用 / Stuck-timer edge instance *)
    tonStuck  : TON;                         (* 卡死判定窗计时器（IN 由变化判据派生 + 相位闸） / Stuck window timer *)
    _bFault   : BOOL;                        (* 故障锁存位 / Latched fault bit *)
    _bCfgBad  : BOOL;                        (* 组态非法当拍量 / Illegal config this scan *)
    _bFin     : BOOL;                        (* 监视值有限性当拍量 / Value finiteness *)
    _bMoved   : BOOL;                        (* 本拍有效变化当拍量（超死区） / Valid move this scan *)
    _bSeen    : BOOL;                        (* 基线已建立标志 / Baseline established flag *)
    _fLast    : REAL;                        (* 基线快照（最近一次有效变化的值）[工程单位] / Baseline snapshot *)
    _fDeltaI  : REAL;                        (* 变化量中间量 [工程单位] / Delta intermediate *)
    _bStuckC  : BOOL;                        (* 卡死起始沿内部单拍量（出口统一映射，R187） / Stuck-edge internal pulse *)
END_VAR
VAR CONSTANT
    DL_SSW_EPS : REAL := 1.0E-6;             (* 判零容差（REAL 量级）[-] / Epsilon *)
END_VAR

(* —— 段 0：当拍判据派生 + 实例无条件刷新（R228A；R_TRIG/TON 全在段 0，无 IF 包裹） —— *)
_bCfgBad := (fDeadband < 0.0) OR NOT (tStuckWin > T#0S);                       (* 死区非负闸 + 卡死窗正域闸 / Deadband and window gates *)
rtReset(CLK := bReset);                                                        (* 复位沿每拍必调 / Reset edge every scan *)
_bFin := (fValue = fValue) AND ((fValue - fValue) = (fValue - fValue));        (* 监视值 NaN 自反 + Inf 差判闸 / Value NaN and Inf gate *)
_fDeltaI := fValue - _fLast;                                                   (* 相对基线变化量（基线无效期不用于判据）[工程单位] / Delta versus baseline *)
_bMoved := _bFin AND _bSeen AND (ABS(_fDeltaI) > fDeadband);                   (* 有效变化：有限 + 基线在 + 超死区（死区 0 即严格不等） / Valid move gate *)
tonStuck(IN := (_eState = E_DL_SswState.eMon) AND _bSeen AND NOT _bMoved AND _bFin, PT := tStuckWin);   (* 卡死窗计时：基线在 + 未变化 + 有限才计时，串 eMon 相位闸 / Stuck timer with phase gate *)
rtStuck(CLK := tonStuck.Q);                                                    (* 卡死窗到点沿每拍必调 / Stuck-elapsed edge every scan *)

(* —— 段 1：单拍量预清零（R107） —— *)
_bStuckC := FALSE;                                                             (* 卡死起始沿内部量预清 / Stuck-edge preset *)
bStuckEdge := FALSE;                                                           (* 卡死起始沿出口预清 / Stuck-edge outlet preset *)
fDelta := 0.0;                                                                 (* 变化量出口预清 / Delta outlet preset *)
fLastMove := T#0S;                                                             (* 最近变化距今出口预清 / Last-move outlet preset *)

(* —— 段 2：复位沿处理（作用域：清故障 + 清报警 + 清基线 + 迁 eIdle，R283 逐项声明） —— *)
IF rtReset.Q THEN
    _bFault := FALSE;                                                          (* 清故障锁存 / Clear fault *)
    _eCause := E_DL_SswCause.eNone;                                            (* 清成因 / Clear cause *)
    bStuck := FALSE;                                                           (* 清卡死报警锁存 / Clear stuck latch *)
    _bSeen := FALSE;                                                           (* 清基线已建立位（重使能重新取基线） / Clear baseline flag *)
    _fLast := 0.0;                                                             (* 清基线快照值 / Clear baseline value *)
    _eState := E_DL_SswState.eIdle;                                            (* 迁未使能相 / Back to idle *)
END_IF

(* —— 段 3：组态故障锁存（锁存至复位沿，R189） —— *)
IF _bCfgBad AND NOT _bFault THEN
    _bFault := TRUE;                                                           (* 锁存故障位 / Latch fault *)
    _eCause := E_DL_SswCause.eCfgIllegal;                                      (* 成因：组态非法 / Cause: illegal config *)
    _eState := E_DL_SswState.eFault;                                           (* 同步迁故障相 / Migrate to fault *)
END_IF

(* —— 段 4：CASE 主状态机（ELSE 兜底迁 eFault，红线 6） —— *)
CASE _eState OF
    E_DL_SswState.eIdle:                                                       (* 未使能：不判死 / Disabled *)
        bStuck := FALSE;                                                       (* 失能清报警出口（eIdle/eFault 出口确定值） / Clear stuck outlet *)
        fDelta := 0.0;                                                         (* 失能清变化量出口 / Clear delta outlet *)
        _bSeen := FALSE;                                                       (* 失能清基线位（重使能重新对齐） / Clear baseline flag *)
        IF bEnable AND NOT _bFault THEN
            _fLast := fValue;                                                  (* 迁入拍取基线首快照（相位闸配套） / Baseline snapshot at entry *)
            _bSeen := TRUE;                                                    (* 基线已建立 / Baseline established *)
            _eState := E_DL_SswState.eMon;                                     (* 使能进入监视 / Enter monitoring *)
        END_IF
    E_DL_SswState.eMon:                                                        (* 监视相：变化刷基线，未变化累计 / Monitoring *)
        IF NOT bEnable THEN
            _eState := E_DL_SswState.eIdle;                                    (* 失能回未使能 / Back to idle *)
        ELSE
            IF _bFin THEN
                fDelta := _fDeltaI;                                            (* 变化量出口（有限拍才派生） / Delta outlet *)
                fLastMove := tonStuck.ET;                                      (* 本窗已积时长镜像 [ms] / Window elapsed mirror *)
            END_IF
            IF _bMoved THEN
                _fLast := fValue;                                              (* 有效变化：基线刷新为当前值（计时器随 IN 翻 FALSE 自动归零） / Refresh baseline on move *)
            END_IF
            IF rtStuck.Q THEN                                                  (* 卡死窗满且全程未变化：报警 / Window elapsed without move *)
                _bStuckC := TRUE;                                              (* 起始沿内部置位（出口统一映射，R187） / Stuck-edge internal *)
                bStuck := TRUE;                                                (* 卡死报警锁存（复位沿清） / Latch stuck alarm *)
                _bFault := TRUE;                                               (* 同步故障锁存（卡死按故障级处理，R45 配对） / Latch fault *)
                _eCause := E_DL_SswCause.eStuck;                               (* 成因：信号卡死（R190 归因唯一） / Cause: signal stuck *)
            END_IF
        END_IF
    E_DL_SswState.eFault:                                                      (* 故障相：冻结保持末值，仅复位沿出 / Fault *)
        ;                                                                      (* 锁存回放（R28） / Replay from latch *)
    ELSE                                                                       (* 非法相位兜底迁安全态 / Illegal phase fallback *)
        _eState := E_DL_SswState.eFault;                                       (* 迁故障相 / To fault *)
        _bFault := TRUE;                                                       (* 同步锁存 / Latch *)
        _eCause := E_DL_SswCause.ePhaseBad;                                    (* 成因：非法相位 / Cause: illegal phase *)
END_CASE

(* —— 段 5：出口映射（内部 _b* → 输出单拍，R187；名实双出口，R191） —— *)
bStuckEdge := _bStuckC;                                                        (* 卡死起始沿单拍出口 / Stuck-edge single-scan outlet *)
bError := _bFault;                                                             (* 故障标志镜像 / Fault flag mirror *)
eState := _eState;                                                             (* 状态出口 / State outlet *)
eCause := _eCause;                                                             (* 成因出口 / Cause outlet *)
END_FUNCTION_BLOCK

(* ---- FB_DL_SimInputBank.st ---- *)
(*
  ==================================================================
  组件名 Component  : FB_DL_SimInputBank
  分类   Category   : DL_Base
  复杂度 Complexity  : cx5
  版本   Version    : 1.0.0
  功能   Purpose    : 调试仿真输入注入组。8 通道手动假值旁路真实输入：通道
                      仿真使能 + 组武装锁存（沿置沿清，防误碰）双闸满足才
                      旁路；退出（通道撤使能 / 组撤武装）自动回真实值；
                      组级与通道级仿真指示出口。与 OutputForcingBank 输出侧
                      强制组成对（R216 互引）。
  来源   Source     : self（库内对称件，R216 互引）
  溯源   Origin     : IEC 61131-3 标准语义的道莅防御性实现；调试输入旁路与
                      武装锁存为公开调试工程语义，clean-room 自研实现，未复
                      制任何厂商私有库源码。
  平台   Platform   : 纯 IEC 61131-3（Standard.library: R_TRIG，无私有库）
  分工声明 Split     : 与 DL_Base 存量 FB_DL_OutputForcingBank 分工——本件为
                      输入侧仿真注入组，OutputForcingBank 为输出侧强制组；
                      本件不做输出强制，也不做信号源切换诊断。
  作者   Author     : 道莅代码库 · PLC 编程专家（R58）
  ------------------------------------------------------------------
  边界 Boundary     :
                      一 双闸条件：组武装 _bArmed（沿锁存）AND 组使能
                         bBankEn AND 通道使能 abSimEn[i]，三者同真才旁路；
                      二 武装锁存解除路径 = bSimDisarmReq 上升沿（唯一沿，
                         R188 头注释声明）；置位路径 = bSimArmReq 上升沿；
                      三 退出自动回真实值：旁路条件任一失效，输出组合逻辑
                         即刻跟随真实输入（无保持延迟）；
                      四 数组按固定界 0..7 遍历（无动态下标，结构性越界
                         防御）；输出 abOut 与输入数组同长度同序；
                      五 无全局变量、无外部变量声明、无物理地址寻址。
  修订记录 Revision  :
    2026-11-21  v1.0.0  R58 首版（批 1 · 序号 2）
  ==================================================================
*)

FUNCTION_BLOCK FB_DL_SimInputBank
VAR_INPUT
    abRealIn     : ARRAY[0..7] OF BOOL; // 真实输入数组（正常过程信号）[-] / the real input array, the normal process signals
    abSimVal     : ARRAY[0..7] OF BOOL; // 仿真假值数组（手动注入）[-] / the simulated value array, manually injected
    abSimEn      : ARRAY[0..7] OF BOOL; // 通道仿真使能数组 [-] / the per channel simulation enable array
    bBankEn      : BOOL := TRUE;  // 组使能（总闸）[-] / the bank enable, the master gate
    bSimArmReq   : BOOL := FALSE; // 武装请求，上升沿置武装锁存 [-] / the arm request, the rising edge raises the arm latch
    bSimDisarmReq: BOOL := FALSE; // 撤武装请求，上升沿清武装锁存 [-] / the disarm request, the rising edge clears the arm latch
END_VAR
VAR_OUTPUT
    abOut      : ARRAY[0..7] OF BOOL; // 混合输出数组（旁路时为假值，否则真实值）[-] / the mixed output array, the fake value when bypassed
    abChnSim   : ARRAY[0..7] OF BOOL; // 通道仿真生效指示数组 [-] / the per channel simulation active array
    bSimActive : BOOL := FALSE; // 组级仿真指示（任一通道旁路中）[-] / the bank simulation indicator, any channel bypassed
    bArmed     : BOOL := FALSE; // 武装锁存指示 [-] / the arm latch indicator
END_VAR
VAR
    rtArm   : R_TRIG; // 武装请求沿检测，段 0 无条件刷新 / the arm request edge, refreshed unconditionally
    rtDisarm: R_TRIG; // 撤武装请求沿检测，段 0 无条件刷新 / the disarm request edge, refreshed unconditionally
    _nI     : DINT;   // 通道遍历索引 [槽] / the channel loop index [slot]
    _bAny   : BOOL;   // 任一通道旁路中工作量 [-] / the any channel bypassed work flag
END_VAR

// 段 0｜沿检测无条件周期刷新（禁入分支）/ segment 0, the unconditional refresh
rtArm(CLK := bSimArmReq); // 武装沿 / the arm edge
rtDisarm(CLK := bSimDisarmReq); // 撤武装沿 / the disarm edge

// 段 1｜武装锁存沿置沿清（边界二，解除路径 = 撤武装上升沿，R188 声明）/ segment 1, the arm latch edge set and edge clear
IF rtArm.Q THEN // 武装上升沿 / the arm rising edge
    bArmed := TRUE; // 置武装锁存 / raise the arm latch
END_IF
IF rtDisarm.Q THEN // 撤武装上升沿（唯一解除路径）/ the disarm rising edge, the only release path
    bArmed := FALSE; // 清武装锁存 / clear the arm latch
END_IF

// 段 2｜通道混合输出（固定界遍历，双闸条件，边界一二三）/ segment 2, the channel mixing, the dual gate
_bAny := FALSE; // 组级指示工作量预置假 / preset the any flag false
FOR _nI := 0 TO 7 DO // 固定界循环，无死循环风险 / the fixed bound loop
    abChnSim[_nI] := bArmed AND bBankEn AND abSimEn[_nI]; // 通道旁路生效判定 / the per channel bypass verdict
    IF abChnSim[_nI] THEN // 旁路生效 / bypassed
        abOut[_nI] := abSimVal[_nI]; // 输出假值 / output the fake value
        _bAny := TRUE; // 组级指示置位 / raise the any flag
    ELSE // 未旁路（边界三：自动回真实值）/ not bypassed, back to the real value
        abOut[_nI] := abRealIn[_nI]; // 输出真实值 / output the real value
    END_IF
END_FOR
bSimActive := _bAny; // 组级仿真指示出口 / the bank simulation indicator
END_FUNCTION_BLOCK

(* ---- FB_DL_SmokeDetZoneMon.st ---- *)
// FB_DL_SmokeDetZoneMon v1.0.0
// 开源溯源：self-cleanroom / 消防域
(*
  道莅工业代码库 | DL_Base | FB_DL_SmokeDetZoneMon
  版本: 1.0.0 | 日期: 2026-11-23 | 轮次: R75
  功能: 消防烟雾探测分区监视：4 分区各自报警/故障/屏蔽三态判定 + 报警
        确认延时去抖 + 报警/故障双锁存（复位沿解除）
  邻件关系: 与 EStopMonitor（急停监视）相邻 —— 差异点：急停件为单点
            安全回路监视，本件为多分区探测三态聚合（报警/故障/屏蔽），
            分区级独立锁存
  锁存声明: 报警锁存 bAnyAlarmLatch 至 bReset 上升沿解除；故障锁存
            bAnyFaultLatch 至该区故障消失且 bReset 上升沿解除（双条件可达）
*)
TYPE E_DL_SmokeZoneState :
(
    eNormal := 0,    // 正常（无报警无故障）/ Normal, no alarm no fault
    eAlarm  := 10,   // 报警（确认延时满）/ Alarm confirmed after delay
    eFault  := 20,   // 探测器故障 / Detector fault
    eMasked := 30     // 分区屏蔽（维护旁路）/ Zone masked for maintenance
);
END_TYPE

FUNCTION_BLOCK FB_DL_SmokeDetZoneMon
VAR_INPUT
    bEnable      : BOOL := FALSE;             // 监视总使能（FALSE 全区置屏蔽态）/ Master enable
    bZoneSmoke1  : BOOL := FALSE;             // 区 1 烟感信号 [-] / Zone 1 smoke signal
    bZoneSmoke2  : BOOL := FALSE;             // 区 2 烟感信号 [-] / Zone 2 smoke signal
    bZoneSmoke3  : BOOL := FALSE;             // 区 3 烟感信号 [-] / Zone 3 smoke signal
    bZoneSmoke4  : BOOL := FALSE;             // 区 4 烟感信号 [-] / Zone 4 smoke signal
    bZoneFault1  : BOOL := FALSE;             // 区 1 探测器故障 [-] / Zone 1 detector fault
    bZoneFault2  : BOOL := FALSE;             // 区 2 探测器故障 [-] / Zone 2 detector fault
    bZoneFault3  : BOOL := FALSE;             // 区 3 探测器故障 [-] / Zone 3 detector fault
    bZoneFault4  : BOOL := FALSE;             // 区 4 探测器故障 [-] / Zone 4 detector fault
    bMask1       : BOOL := FALSE;             // 区 1 屏蔽请求 [-] / Zone 1 mask request
    bMask2       : BOOL := FALSE;             // 区 2 屏蔽请求 [-] / Zone 2 mask request
    bMask3       : BOOL := FALSE;             // 区 3 屏蔽请求 [-] / Zone 3 mask request
    bMask4       : BOOL := FALSE;             // 区 4 屏蔽请求 [-] / Zone 4 mask request
    tAlarmDelay  : TIME := T#5S;              // 报警确认延时 [ms]，去抖 / Alarm confirm delay
    bReset       : BOOL := FALSE;             // 复位（上升沿解锁存）/ Reset, rising edge clears latches
END_VAR
VAR_OUTPUT
    eState1          : E_DL_SmokeZoneState;   // 区 1 三态 / Zone 1 state
    eState2          : E_DL_SmokeZoneState;   // 区 2 三态 / Zone 2 state
    eState3          : E_DL_SmokeZoneState;   // 区 3 三态 / Zone 3 state
    eState4          : E_DL_SmokeZoneState;   // 区 4 三态 / Zone 4 state
    bAnyAlarmLatch   : BOOL;                  // 任一区报警锁存（复位沿解除）/ Any alarm latched
    bAnyFaultLatch   : BOOL;                  // 任一区故障锁存 / Any fault latched
    uAlarmZoneCnt    : UDINT;                 // 当前报警区数 [区] / Current alarm zone count
    uFaultZoneCnt    : UDINT;                 // 当前故障区数 [区] / Current fault zone count
    bValid           : BOOL;                  // 组态有效回执 [-] / Config validity receipt
    bError           : BOOL;                  // 故障标志（延时组态非法）/ Fault flag (delay config illegal)
    uErrorId         : UDINT;                 // 事件码，0 = 无事件；16#0002_2401 = 延时组态非法 / Event code
END_VAR
VAR
    rtrReset     : R_TRIG;                    // 复位沿（每拍无条件刷新）/ Reset edge, refreshed every cycle
    tonZone1     : TON;                       // 区 1 确认延时（自复位）/ Zone 1 confirm delay, self-resetting
    tonZone2     : TON;                       // 区 2 确认延时 / Zone 2 confirm delay
    tonZone3     : TON;                       // 区 3 确认延时 / Zone 3 confirm delay
    tonZone4     : TON;                       // 区 4 确认延时 / Zone 4 confirm delay
    bLatch1      : BOOL;                      // 区 1 报警锁存 [-] / Zone 1 alarm latch
    bLatch2      : BOOL;                      // 区 2 报警锁存 [-] / Zone 2 alarm latch
    bLatch3      : BOOL;                      // 区 3 报警锁存 [-] / Zone 3 alarm latch
    bLatch4      : BOOL;                      // 区 4 报警锁存 [-] / Zone 4 alarm latch
    bFltLatch1   : BOOL;                      // 区 1 故障锁存 [-] / Zone 1 fault latch
    bFltLatch2   : BOOL;                      // 区 2 故障锁存 [-] / Zone 2 fault latch
    bFltLatch3   : BOOL;                      // 区 3 故障锁存 [-] / Zone 3 fault latch
    bFltLatch4   : BOOL;                      // 区 4 故障锁存 [-] / Zone 4 fault latch
END_VAR

// —— 段 0：实例无条件刷新（R7：沿与定时器每周期调用） —— //
rtrReset(CLK := bReset);                          // 复位沿每拍刷新 / Reset edge refreshed
tonZone1(IN := bEnable AND bZoneSmoke1 AND (NOT bMask1), PT := tAlarmDelay);   // 区 1 延时 / Zone 1 delay
tonZone2(IN := bEnable AND bZoneSmoke2 AND (NOT bMask2), PT := tAlarmDelay);   // 区 2 延时 / Zone 2 delay
tonZone3(IN := bEnable AND bZoneSmoke3 AND (NOT bMask3), PT := tAlarmDelay);   // 区 3 延时 / Zone 3 delay
tonZone4(IN := bEnable AND bZoneSmoke4 AND (NOT bMask4), PT := tAlarmDelay);   // 区 4 延时 / Zone 4 delay

// —— 段 1：组态闸 —— //
bValid := (tAlarmDelay > T#0MS);                  // 延时必须非零（去抖有效）/ Delay must be nonzero
IF NOT bValid THEN
    bError   := TRUE;                             // 故障级：延时组态非法 / Fault level: delay config illegal
    uErrorId := 16#0002_2401;                     // 故障码（24xx 步进）/ Fault code
    RETURN;                                       // 非法组态不判定 / No judgment on illegal config
END_IF
bError   := FALSE;                                // 组态恢复：故障清零（解除路径）/ Fault cleared on valid config
uErrorId := 16#0000;                              // 事件码清零 / Event code cleared

// —— 段 2：复位沿解锁存（双条件可达：锁存源消失 + 复位沿） —— //
IF rtrReset.Q THEN
    IF NOT bZoneSmoke1 THEN
        bLatch1 := FALSE;                         // 区 1 报警锁存解除 / Zone 1 alarm latch clear
    END_IF
    IF NOT bZoneSmoke2 THEN
        bLatch2 := FALSE;                         // 区 2 报警锁存解除 / Zone 2 clear
    END_IF
    IF NOT bZoneSmoke3 THEN
        bLatch3 := FALSE;                         // 区 3 报警锁存解除 / Zone 3 clear
    END_IF
    IF NOT bZoneSmoke4 THEN
        bLatch4 := FALSE;                         // 区 4 报警锁存解除 / Zone 4 clear
    END_IF
    IF NOT bZoneFault1 THEN
        bFltLatch1 := FALSE;                      // 区 1 故障锁存解除 / Zone 1 fault clear
    END_IF
    IF NOT bZoneFault2 THEN
        bFltLatch2 := FALSE;                      // 区 2 故障锁存解除 / Zone 2 clear
    END_IF
    IF NOT bZoneFault3 THEN
        bFltLatch3 := FALSE;                      // 区 3 故障锁存解除 / Zone 3 clear
    END_IF
    IF NOT bZoneFault4 THEN
        bFltLatch4 := FALSE;                      // 区 4 故障锁存解除 / Zone 4 clear
    END_IF
END_IF

// —— 段 3：报警/故障锁存置位（源出现即置位，状态型锁存） —— //
IF bEnable AND (NOT bMask1) THEN
    IF tonZone1.Q THEN
        bLatch1 := TRUE;                          // 确认延时满：区 1 报警锁存 / Delay full: zone 1 alarm latch
    END_IF
END_IF
IF bEnable AND (NOT bMask2) THEN
    IF tonZone2.Q THEN
        bLatch2 := TRUE;                          // 区 2 报警锁存 / Zone 2 alarm latch
    END_IF
END_IF
IF bEnable AND (NOT bMask3) THEN
    IF tonZone3.Q THEN
        bLatch3 := TRUE;                          // 区 3 报警锁存 / Zone 3 alarm latch
    END_IF
END_IF
IF bEnable AND (NOT bMask4) THEN
    IF tonZone4.Q THEN
        bLatch4 := TRUE;                          // 区 4 报警锁存 / Zone 4 alarm latch
    END_IF
END_IF
IF bEnable AND bZoneFault1 AND (NOT bMask1) THEN
    bFltLatch1 := TRUE;                           // 区 1 故障锁存 / Zone 1 fault latch
END_IF
IF bEnable AND bZoneFault2 AND (NOT bMask2) THEN
    bFltLatch2 := TRUE;                           // 区 2 故障锁存 / Zone 2 fault latch
END_IF
IF bEnable AND bZoneFault3 AND (NOT bMask3) THEN
    bFltLatch3 := TRUE;                           // 区 3 故障锁存 / Zone 3 fault latch
END_IF
IF bEnable AND bZoneFault4 AND (NOT bMask4) THEN
    bFltLatch4 := TRUE;                           // 区 4 故障锁存 / Zone 4 fault latch
END_IF

// —— 段 4：逐区三态判定（故障 > 报警 > 屏蔽 > 正常优先序） —— //
IF (NOT bEnable) OR bMask1 THEN
    eState1 := E_DL_SmokeZoneState.eMasked;       // 区 1 屏蔽（失能按屏蔽安全语义）/ Zone 1 masked
ELSIF bFltLatch1 THEN
    eState1 := E_DL_SmokeZoneState.eFault;        // 区 1 故障 / Zone 1 fault
ELSIF bLatch1 THEN
    eState1 := E_DL_SmokeZoneState.eAlarm;        // 区 1 报警 / Zone 1 alarm
ELSE
    eState1 := E_DL_SmokeZoneState.eNormal;       // 区 1 正常 / Zone 1 normal
END_IF
IF (NOT bEnable) OR bMask2 THEN
    eState2 := E_DL_SmokeZoneState.eMasked;       // 区 2 屏蔽 / Zone 2 masked
ELSIF bFltLatch2 THEN
    eState2 := E_DL_SmokeZoneState.eFault;        // 区 2 故障 / Zone 2 fault
ELSIF bLatch2 THEN
    eState2 := E_DL_SmokeZoneState.eAlarm;        // 区 2 报警 / Zone 2 alarm
ELSE
    eState2 := E_DL_SmokeZoneState.eNormal;       // 区 2 正常 / Zone 2 normal
END_IF
IF (NOT bEnable) OR bMask3 THEN
    eState3 := E_DL_SmokeZoneState.eMasked;       // 区 3 屏蔽 / Zone 3 masked
ELSIF bFltLatch3 THEN
    eState3 := E_DL_SmokeZoneState.eFault;        // 区 3 故障 / Zone 3 fault
ELSIF bLatch3 THEN
    eState3 := E_DL_SmokeZoneState.eAlarm;        // 区 3 报警 / Zone 3 alarm
ELSE
    eState3 := E_DL_SmokeZoneState.eNormal;       // 区 3 正常 / Zone 3 normal
END_IF
IF (NOT bEnable) OR bMask4 THEN
    eState4 := E_DL_SmokeZoneState.eMasked;       // 区 4 屏蔽 / Zone 4 masked
ELSIF bFltLatch4 THEN
    eState4 := E_DL_SmokeZoneState.eFault;        // 区 4 故障 / Zone 4 fault
ELSIF bLatch4 THEN
    eState4 := E_DL_SmokeZoneState.eAlarm;        // 区 4 报警 / Zone 4 alarm
ELSE
    eState4 := E_DL_SmokeZoneState.eNormal;       // 区 4 正常 / Zone 4 normal
END_IF

// —— 段 5：聚合输出（计数用枚举统计，锁存聚合） —— //
uAlarmZoneCnt := 0;                               // 报警区计数预清 / Alarm zone count preset
IF eState1 = E_DL_SmokeZoneState.eAlarm THEN
    uAlarmZoneCnt := uAlarmZoneCnt + 1;           // 区 1 计入 / Zone 1 counted
END_IF
IF eState2 = E_DL_SmokeZoneState.eAlarm THEN
    uAlarmZoneCnt := uAlarmZoneCnt + 1;           // 区 2 计入 / Zone 2 counted
END_IF
IF eState3 = E_DL_SmokeZoneState.eAlarm THEN
    uAlarmZoneCnt := uAlarmZoneCnt + 1;           // 区 3 计入 / Zone 3 counted
END_IF
IF eState4 = E_DL_SmokeZoneState.eAlarm THEN
    uAlarmZoneCnt := uAlarmZoneCnt + 1;           // 区 4 计入 / Zone 4 counted
END_IF
uFaultZoneCnt := 0;                               // 故障区计数预清 / Fault zone count preset
IF eState1 = E_DL_SmokeZoneState.eFault THEN
    uFaultZoneCnt := uFaultZoneCnt + 1;           // 区 1 计入 / Zone 1 counted
END_IF
IF eState2 = E_DL_SmokeZoneState.eFault THEN
    uFaultZoneCnt := uFaultZoneCnt + 1;           // 区 2 计入 / Zone 2 counted
END_IF
IF eState3 = E_DL_SmokeZoneState.eFault THEN
    uFaultZoneCnt := uFaultZoneCnt + 1;           // 区 3 计入 / Zone 3 counted
END_IF
IF eState4 = E_DL_SmokeZoneState.eFault THEN
    uFaultZoneCnt := uFaultZoneCnt + 1;           // 区 4 计入 / Zone 4 counted
END_IF
bAnyAlarmLatch := (uAlarmZoneCnt > 0);            // 任一报警聚合（当前态镜像）/ Any alarm aggregate
bAnyFaultLatch := (uFaultZoneCnt > 0);            // 任一故障聚合 / Any fault aggregate
END_FUNCTION_BLOCK

(* ---- FB_DL_SRBistable.st ---- *)
(*==============================================================================
 * 组件名称 (Component)  : FB_DL_SRBistable
 * 所属子库 (Sublibrary) : DL_Base
 * 当前版本 (Version)    : 1.0.0
 * 兼容性   (Platform)   : CODESYS 3.5 / TwinCAT 3 / 汇川 InoProShop / Machine Expert
 *                         仅依赖纯 IEC 61131-3 标准运算符，零厂商方言
 * 功能描述 (Function)   : SR 置位优先双稳态防御包装。内部委托 IEC 61131-3 标准
 *                         SR 语义（bQ1 := bS1 OR (bQ1 AND NOT bR)），外围提供
 *                         S1/R 同拍仲裁显式化与仲裁诊断码输出。
 * 溯源     (Origin)     : IEC 61131-3 标准语义的道莅防御性实现
 *                         （接口语义由 IEC 61131-3 定义，clean-room 重写，
 *                         参考公开标准条款）
 * 码位     (Diag Codes) : 信息级占用区间 16#0001_014D（本件独占，仅此一码）
 *                         16#0001_014D = S1/R 同拍为 TRUE，置位胜出（标准语义，
 *                         仅供现场排查，不置故障）
 * 类型裁定 (Type Note)  : 码位段 16#0001_xxxx 为全库共享 32 位段，WORD 容量不足，
 *                         故 uDiag 采用 UDINT 承载（与库内 uErrorId : UDINT 惯例一致）
 * 依赖     (Depends)    : 无 DL_ 内部依赖；无标准库实例（纯布尔逻辑）
 * 红线自检 (Redline)    : R1 ✓ 零全局变量与外部变量引用 ｜ R2 ✓ 零物理 IO 地址直写
 *                         R3 ✓ 纯 IEC 61131-3 ｜ R4 ✓ 同拍仲裁显式化+首扫初始化
 *                         R5 ✓ 全变量中英双语同行注释 ｜ R6 N/A（无顺序状态机，见下）
 *                         R7 ✓ 无定时器/沿检测实例（N/A）
 * 说明     (Note)       : R6 标注 N/A —— 本组件为组合逻辑双稳态，不存在顺序状态机，
 *                         无 CASE 可写；非法状态不可能出现（唯一状态即输出锁存），
 *                         故以本节说明替代 ELSE 兜底，符合"无状态机则标注 N/A"口径。
 * 防御行为声明 (Defense): ① S1 与 R 同拍为 TRUE 时按 IEC 语义置位优先（S1 胜出），
 *                           同时置信息级诊断码 16#0001_014D，下拍仲裁消失自动清零；
 *                         ② 首扫输出初始化为 FALSE，杜绝上电假输出。
 * 修订历史 (Revision)   :
 *   2026-11-16  v1.0.0  首版入库（R14 批 1 · T0 快车道）
 *============================================================================*)
FUNCTION_BLOCK FB_DL_SRBistable
VAR_INPUT
    bS1 : BOOL;  // 置位主导输入（IEC S1 语义），TRUE 时输出无条件置位 / Set-dominant input (IEC S1), TRUE forces output set
    bR  : BOOL;  // 复位输入，仅在 S1 为 FALSE 的拍次生效 / Reset input, effective only on scans where S1 is FALSE
END_VAR
VAR_OUTPUT
    bQ1   : BOOL;   // 置位优先输出（IEC Q1 语义），TRUE 保持至复位 / Set-dominant output (IEC Q1), latched TRUE until reset
    uDiag : UDINT;  // 仲裁诊断字，16#0001_014D=S1/R 同拍置位胜出，0=无仲裁事件 / Arbitration diag word, 16#0001_014D=same-scan S1/R with set winning, 0=no arbitration
END_VAR
VAR
    xInit : BOOL;   // 首扫初始化标志，FALSE=尚未完成上电初始化 / First-scan init flag, FALSE = power-on init not yet done
END_VAR

(*------------------------------------------------------------------------------
 * 段 1｜首扫初始化（历史教训⑤口径）：置于逻辑最前，禁止"初值置位后同步清零"反模式
 *      First-scan init (lesson 5): placed at the very front of the logic body
 *-----------------------------------------------------------------------------*)
IF NOT xInit THEN
    xInit := TRUE;      // 置初始化完成标志 / Mark init as done
    bQ1   := FALSE;     // 首扫输出强制 FALSE，杜绝上电假输出 / Force output FALSE on first scan
    uDiag := 16#0000_0000;  // 首扫诊断字清零 / Clear diag word on first scan
END_IF

(*------------------------------------------------------------------------------
 * 段 2｜同拍仲裁诊断：S1 与 R 同拍为 TRUE 是标准定义的合法竞态，置信息码不置故障
 *      Same-scan arbitration diag: S1 AND R is a legal race per the standard,
 *      informational code only, never a fault
 *-----------------------------------------------------------------------------*)
IF bS1 AND bR THEN
    uDiag := 16#0001_014D;  // 同拍竞态：置位优先胜出（信息级）/ Same-scan race: set-dominant wins (informational)
ELSE
    uDiag := 16#0000_0000;  // 无竞态，诊断字清零 / No race, clear diag word
END_IF

(*------------------------------------------------------------------------------
 * 段 3｜SR 置位优先核心语义（委托 IEC 61131-3 标准 SR 定义，不重实现）：
 *      bQ1 := bS1 OR (bQ1 AND NOT bR)，右侧 bQ1 取上一拍锁存值
 *      SR set-dominant core semantics (delegates to the IEC 61131-3 SR definition);
 *      the bQ1 on the right-hand side reads the latched value of the previous scan
 *-----------------------------------------------------------------------------*)
bQ1 := bS1 OR (bQ1 AND NOT bR);  // 置位优先：S1=1 恒置位，S1=0 且 R=1 才复位 / Set-dominant: S1=1 always sets, reset only when S1=0 and R=1
END_FUNCTION_BLOCK

(* ---- FB_DL_SrEx.st ---- *)
(*==============================================================================
 * 组件名称 (Component)  : FB_DL_SrEx
 * 所属子库 (Sublibrary) : DL_Base
 * 当前版本 (Version)    : 1.0.0
 * 兼容性   (Platform)   : CODESYS 3.5 / TwinCAT 3 / 汇川 InoProShop / Machine Expert
 *                         仅依赖纯 IEC 61131-3 标准运算符，零厂商方言
 * 功能描述 (Function)   : SR 置位优先双稳态防御包装。内部委托 IEC 61131-3 标准
 *                         SR 语义（bQ1 := bS1 OR (bQ1 AND NOT bR)），外围提供
 *                         S1/R 同拍仲裁显式化诊断与主从双输出镜像。
 * 溯源     (Origin)     : IEC 61131-3 标准语义的道莅防御性实现
 *                         （接口语义由 IEC 61131-3 定义，clean-room 重写，
 *                         参考公开标准条款，未复制任何闭源厂商源码）
 * 码位     (Diag Codes) : 信息级占用区间 16#0001_049A（本件独占，仅此一码）
 *                         16#0001_049A = S1/R 同拍为 TRUE，置位胜出（标准语义，
 *                         仅供现场排查，不置故障）
 *                         （R90 反证句：同拍仲裁事实无法由 bQ1 观测——置位胜出与
 *                           单纯置位的输出同为 TRUE，现有输出组合无法还原「曾发生
 *                           同拍竞争」，故占信息码）
 * 类型裁定 (Type Note)  : 码位段 16#0001_xxxx 为全库共享 32 位段，WORD 容量不足，
 *                         故 uDiag 采用 UDINT 承载（与库内 uErrorId : UDINT 惯例一致）
 * 依赖     (Depends)    : 无 DL_ 内部依赖；无标准库实例（纯布尔逻辑）
 * 红线自检 (Redline)    : R1 ✓ 零全局变量与外部变量引用 ｜ R2 ✓ 零物理 IO 地址直写
 *                         R3 ✓ 纯 IEC 61131-3 ｜ R4 ✓ 同拍仲裁显式化，无浮点无除法
 *                         R5 ✓ 全变量中英双语同行注释 ｜ R6 N/A（无顺序状态机，见下）
 *                         R7 N/A 无定时器与沿检测实例（纯组合保持逻辑）
 * 说明     (Note)       : R6 标注 N/A —— 本组件为单步双稳态保持逻辑，不存在顺序
 *                         状态机，无 CASE 可写；非法状态不可能出现（唯一状态即
 *                         「保持 / 置位 / 复位」三态组合，由标准布尔语义全覆盖），
 *                         故以本节说明替代 ELSE 兜底，符合"无状态机则标注 N/A"口径。
 * 输出语义声明 (R191)   : bS1 = FALSE 且 bR = FALSE 时输出保持末值（双稳态记忆语义），
 *                         非降级非冻结，由标准 SR 语义保证；主从输出 bQ1 与 bQ1M
 *                         单点同源赋值（名实双出口，R191 名实相符）。
 * 修订历史 (Revision)   :
 *   2026-11-19  v1.0.0  首版入库（R40 批 4 · T0 快车道）
 *============================================================================*)
FUNCTION_BLOCK FB_DL_SrEx
VAR_INPUT
    bS1 : BOOL; // 置位输入，TRUE 请求置位，与复位同拍时置位优先胜出 ｜ set input, TRUE requests set, wins the arbitration when simultaneous with the reset
    bR  : BOOL; // 复位输入，TRUE 请求复位，与置位同拍时被置位优先压制 ｜ reset input, TRUE requests reset, suppressed when simultaneous with the set
END_VAR
VAR_OUTPUT
    bQ1   : BOOL;  // 主输出，置位优先双稳态 ｜ main output of the set-dominant bistable
    bQ1M  : BOOL;  // 从输出，与 bQ1 同源镜像（名实双出口）｜ mirror output, same source as bQ1
    uDiag : UDINT; // 诊断字，16#0001_049A=S1/R 同拍置位胜出，0=无诊断事件 ｜ diag word, 16#0001_049A=set wins on simultaneous S1/R, 0=no diag event
END_VAR

// 段 1｜SR 置位优先标准语义主体（IEC 61131-3 双稳态，不重实现状态内核） ｜ SR set-dominant standard semantics (IEC 61131-3 bistable, no kernel re-implementation)
bQ1 := bS1 OR (bQ1 AND NOT bR); // 置位优先：S1 为真置位，R 单独为真复位，同拍置位胜出 ｜ set-dominant: S1 sets, R alone resets, the set wins on simultaneity

// 段 2｜同拍仲裁显式化诊断（信息级每拍重算口径） ｜ simultaneous-arbitration diagnostics (info level, recomputed every scan)
IF bS1 AND bR THEN
    uDiag := 16#0001_049A; // 同拍仲裁：置位优先胜出（信息级，仅排查用）｜ simultaneous arbitration: the set wins (info level, for troubleshooting only)
ELSE
    uDiag := 16#0000_0000; // 无同拍仲裁事件，清码（信息级允许每拍重算）｜ no arbitration event, clear the code (info level may be recomputed per scan)
END_IF

// 段 3｜主从输出镜像：单点同源赋值（R191 名实双出口） ｜ main-mirror output: single same-source assignment (R191 paired exits)
bQ1M := bQ1; // 从输出镜像主输出 ｜ the mirror output copies the main output
END_FUNCTION_BLOCK

(* ---- FB_DL_StepSequencer.st ---- *)
(*==============================================================================
 * 组件名称 (Component)  : FB_DL_StepSequencer
 * 所属子库 (Sublibrary) : DL_Base
 * 当前版本 (Version)    : 1.0.1
 * 兼容性   (Platform)   : CODESYS 3.5 / TwinCAT 3 / 汇川 InoProShop / Machine Expert
 *                         仅依赖 Standard.library（TON / R_TRIG），零厂商方言
 * 功能描述 (Function)   : 通用顺控步引擎（顺序功能图的 ST 基类形态）。
 *                         只管理"当前步号、步内计时、步超时、推进、暂停、单步、故障锁存"，
 *                         动作不写死在块内：调用方按当前步号执行动作，并按步号回报完成信号。
 *                         因此本块可作为上百个工站的共用基类，而不是某个工站的专用代码。
 *                         每步可配独立超时，超时锁定故障并记录故障步号，便于现场定位；
 *                         步完成信号为电平语义，换步后第一个周期屏蔽完成判定，
 *                         从结构上杜绝"旧步残留完成位导致连环跳步"的不稳定转换。
 * 开源溯源 (Origin)     : 原创实现。步状态机与步超时监控为顺序功能图最佳实践的公开共识；
 *                         通用步引擎的职责切分（动作外置）为本库差异化设计，未复制任何源码。
 * 本文件内含       : TYPE  E_DL_SeqState（配套枚举，归属 DL_Base）
 *                    FB    FB_DL_StepSequencer
 * 依赖     (Depends)    : 无 DL_ 内部依赖；Standard.library: TON / R_TRIG
 * 红线自检 (Redline)    : R1 ✓ 禁用全局存储与物理寻址 ｜ R2 ✓ 无地址直写
 *                         R3 ✓ 纯 IEC 61131-3 ｜ R4 ✓ 步号双检 + 超时钳位 + 非法状态兜底
 *                         R5 ✓ 全变量中英双语同行注释 ｜ R6 ✓ 五态 ENUM + CASE + ELSE 兜底
 *                         R7 ✓ 五个实例主体最前部无条件刷新（本组件核心考点）
 *                         R8 ✓ 步数与超时上限全常量化
 *
 * 【完成信号电平语义 / Level-semantic step-done signals（决策 D-R2-09，边界 B12）】
 *   调用方在当前步的条件满足时把对应位保持 TRUE，顺控器在推进瞬间屏蔽该位一个周期。
 *   调用方必须在新步开始后撤销旧步的完成位：本块只屏蔽一个周期，
 *   若旧位长期保持 TRUE 且新步恰好也读该索引，仍会被判成立。
 *   Callers must drop the previous step's done bit once the step has advanced.
 *
 * 【暂停语义 / Hold semantics（决策 D-R2-10，边界 B5）】
 *   暂停期间步计时冻结（定时器输入断开，已计时清零），恢复后**重新计时**而不是续算。
 *   "暂停续算"需要差分补偿，会让定时器语义复杂化；代价是本块明确披露"暂停不算超时"。
 *
 * 【单步调试 / Single-step commissioning（边界 B6）】
 *   单步模式下每步完成即进入暂停态，等待推进沿才真正换步，供维护工程师逐段验证。
 *
 * 【断电保持 / Retain（边界 B12）】
 *   是否将实例声明为断电保持由调用方按工艺决定：保持可续跑，不保持则复位到空闲。
 *
 * 修订历史 (Revision)   :
 *   2026-11-14  v1.0.0  首版入库（Phase 1 第二轮 · Level 0 批次 D）
 *   2026-11-14  v1.0.1  修复故障码不锁存缺陷：原实现在每周期开头无条件清零 uErrorId，
 *                       而故障态分支不再重写故障码，导致进入故障后的下一个扫描周期
 *                       bError 仍为 TRUE、uErrorId 却读回 0，现场与 HMI 丢失根因。
 *                       改为故障锁存期间保留进入故障时的故障码，仅复位沿清零。
 *============================================================================*)

(*-----------------------------------------------------------------------------
 * 枚举: E_DL_SeqState（归属 DL_Base，与 FB_DL_StepSequencer 同文件）
 * 含义: 顺控引擎主状态。数值步长留空位便于后续插态而不破坏已有工程。
 *----------------------------------------------------------------------------*)
TYPE E_DL_SeqState :
(
    eIdle  := 0,     // 空闲待机：步号无效，等待启动沿 / Idle, no active step, waiting for the start edge
    eRun   := 10,    // 运行中：执行当前步动作并监控完成与超时 / Running, executing the current step
    eHold  := 20,    // 暂停：单步调试等待推进沿 / Held, single-step mode waiting for the advance edge
    eDone  := 30,    // 全部步完成：步号保持末步 / All steps done, the step index holds the last step
    eFault := 99     // 故障锁定：步超时或非法状态，仅复位沿可解除 / Fault latched, only the reset edge clears it
);
END_TYPE

FUNCTION_BLOCK FB_DL_StepSequencer
VAR_INPUT
    bStart        : BOOL;                       // 上升沿：从 0 号步启动 / Rising edge: start from step 0
    abStepDone    : ARRAY[0..15] OF BOOL;       // 步完成信号（电平，调用方按当前步维护）/ Step-done levels, caller-maintained
    auStepTimeout : ARRAY[0..15] OF TIME;       // 每步超时 [ms]，0 = 该步不监控 / Per-step timeout [ms], 0 = not monitored
    bHold         : BOOL := FALSE;              // TRUE = 暂停：冻结推进与超时计时 / TRUE = hold advancing and the timeout
    bSingleStep   : BOOL := FALSE;              // TRUE = 单步调试模式 / Single-step commissioning mode
    bAdvance      : BOOL;                       // 单步模式下上升沿推进一步 / Rising edge: advance one step in single-step mode
    bAbort        : BOOL;                       // 上升沿：中止回空闲，不设故障码 / Rising edge: abort to idle without an error
    bReset        : BOOL;                       // 上升沿：清除故障回空闲 / Rising edge: clear the fault and return to idle
END_VAR
VAR_OUTPUT
    nCurrentStep  : INT;     // 当前步号 0..15，-1 = 未运行 / Current step 0..15, -1 = inactive
    bRunning      : BOOL;    // 运行状态标志 / Running flag
    bDone         : BOOL;    // 全部步完成 / All steps done
    bError        : BOOL;    // 故障标志，bReset 清除 / Fault flag, cleared by bReset
    nFaultStep    : INT;     // 超时故障发生步号，-1 = 无 / Fault step index, -1 = none
    tStepElapsed  : TIME;    // 当前步已运行时间 [ms] / Elapsed time in the current step [ms]
    uErrorId      : UDINT;   // 故障码，0 = 无故障 / Error code, 0 = no error
END_VAR
VAR
    eState        : E_DL_SeqState;   // 主状态机 / Main state machine
    fbTonStep     : TON;             // 步计时器 / Step timer
    fbTrigStart   : R_TRIG;          // 启动沿检测实例 / Start edge detector instance
    fbTrigAbort   : R_TRIG;          // 中止沿检测实例 / Abort edge detector instance
    fbTrigReset   : R_TRIG;          // 复位沿检测实例 / Reset edge detector instance
    fbTrigAdvance : R_TRIG;          // 单步推进沿检测实例 / Advance edge detector instance
    nStep         : INT;             // 内部步号 / Internal step index
    tEffTimeout   : TIME;            // 当前步生效超时（已钳位）[ms] / Clamped effective timeout of the current step [ms]
    bTimeoutArmed : BOOL;            // 当前步是否启用超时监控 / Timeout monitoring armed for the current step
    bJustAdvanced : BOOL;            // 换步后首周期屏蔽标志（按下一拍提交）/ First-scan-after-advance mask, committed one scan later
    bMaskNext     : BOOL;            // 下一周期屏蔽请求 / Mask request for the next scan
    bDoAdvance    : BOOL;            // 本周期请求推进 / Advance requested this scan
    bArmStep      : BOOL;            // 本周期请求装载步超时 / Step timeout load requested this scan
    bSkipSm       : BOOL;            // 本周期跳过状态机（复位 / 中止已处理）/ Skip the state machine this scan
    bFirstScan    : BOOL := TRUE;    // 上电首扫初始化标志 / First-scan initialisation flag
END_VAR
VAR CONSTANT
    DL_SEQ_MAX_STEPS : INT  := 16;      // 步数上限 [步]，与数组维度一致 / Step count, must match the arrays
    DL_SEQ_IDX_NONE  : INT  := -1;      // 无效步号哨兵 / Sentinel for no step
    DL_SEQ_TOUT_MAX  : TIME := T#12H;   // 单步超时上限钳位 [ms] / Per-step timeout clamp [ms]
END_VAR

(*------------------------------------------------------------------------------
 * 段 1｜无条件刷新区（红线 R7 / 边界 B1）：四沿 + 一步计时，全部位于主体最前部
 *      Unconditional refresh zone: four edge instances plus the step timer
 *      IN 由"状态 + 暂停 + 超时启用 + 换步屏蔽"先行推导成 BOOL，实例调用本身无条件
 *      IN is derived into a BOOL first, the instance call itself stays unconditional
 *-----------------------------------------------------------------------------*)
fbTrigStart(CLK   := bStart);
fbTrigAbort(CLK   := bAbort);
fbTrigReset(CLK   := bReset);
fbTrigAdvance(CLK := bAdvance);

fbTonStep(IN := (eState = eRun) AND (NOT bHold) AND bTimeoutArmed AND (NOT bJustAdvanced),
          PT := tEffTimeout);

(*------------------------------------------------------------------------------
 * 段 2｜上电首扫初始化：步号与故障步号必须显式置为无效哨兵，不能依赖默认零
 *      First-scan init: step indices must be set to the sentinel, never left at zero
 *-----------------------------------------------------------------------------*)
IF bFirstScan THEN
    bFirstScan := FALSE;
    eState     := eIdle;
    nStep      := DL_SEQ_IDX_NONE;
    nFaultStep := DL_SEQ_IDX_NONE;
END_IF

(*------------------------------------------------------------------------------
 * 段 3｜故障码清零口径（v1.0.1 修正）：故障锁存期间必须保留进入故障时的故障码
 *      Error-code policy: while the fault is latched the entry code must survive
 *      故障码是"锁存事实"而非"本周期瞬时量"：若每周期无条件清零，
 *      进入故障后的下一拍就会读回 0，HMI 与现场工程师同时丢失根因
 *      A fault code is a latched fact; an unconditional clear would erase it one scan later
 *-----------------------------------------------------------------------------*)
IF eState <> eFault THEN
    uErrorId := 16#0000_0000;
END_IF

(*------------------------------------------------------------------------------
 * 段 4｜复位与中止（边界 B7/B9）：复位仅在故障态有效，中止在非故障态有效
 *      Reset works only in fault, abort works everywhere except fault
 *      两者都清空步号与计时，中止刻意不设故障码——操作员主动中止不是故障
 *      Abort raises no error because a deliberate operator stop is not a fault
 *-----------------------------------------------------------------------------*)
bSkipSm    := FALSE;
bDoAdvance := FALSE;
bArmStep   := FALSE;

IF fbTrigReset.Q AND (eState = eFault) THEN
    eState        := eIdle;
    nStep         := DL_SEQ_IDX_NONE;
    nFaultStep    := DL_SEQ_IDX_NONE;
    tEffTimeout   := T#0S;
    bTimeoutArmed := FALSE;
    uErrorId      := 16#0000_0000;   // 故障码唯一清除路径 / The only path that clears the fault code
    bMaskNext     := TRUE;
    bSkipSm       := TRUE;
END_IF

IF fbTrigAbort.Q AND (eState <> eFault) THEN
    eState        := eIdle;
    nStep         := DL_SEQ_IDX_NONE;
    tEffTimeout   := T#0S;
    bTimeoutArmed := FALSE;
    bMaskNext     := TRUE;
    bSkipSm       := TRUE;
END_IF

(*------------------------------------------------------------------------------
 * 段 5｜主状态机（红线 R6 / 边界 B10）：ENUM + CASE + ELSE 兜底
 *      Main state machine with the mandatory ELSE fallback
 *-----------------------------------------------------------------------------*)
IF NOT bSkipSm THEN

    CASE eState OF

        eIdle:
            (* 启动沿：从 0 号步开始，并装载该步超时 *)
            (* Start edge: begin at step 0 and load its timeout *)
            IF fbTrigStart.Q THEN
                nStep         := 0;
                bArmStep      := TRUE;
                bMaskNext     := TRUE;
                eState        := eRun;
            END_IF

        eRun:
            (*------------------------------------------------------------------
             * 段 5a｜超时优先（边界 B4）：先判超时再判完成，避免"超时同时完成"时漏报
             *      Timeout first: a timeout wins over a simultaneous completion
             *-----------------------------------------------------------------*)
            IF fbTonStep.Q THEN
                eState     := eFault;
                nFaultStep := nStep;
                uErrorId   := 16#0001_000B;
            ELSIF (NOT bHold) AND (NOT bJustAdvanced) THEN

                (*--------------------------------------------------------------
                 * 段 5b｜完成判定（边界 B2/B11）：只采当前步，且换步首周期不采
                 *      Completion: only the current step, never in the first scan after a switch
                 *-------------------------------------------------------------*)
                IF (nStep >= 0) AND (nStep < DL_SEQ_MAX_STEPS) THEN
                    IF abStepDone[nStep] THEN
                        IF bSingleStep THEN
                            (* 单步模式：完成即暂停，等推进沿再换步 *)
                            (* Single-step: hold after completion until the advance edge *)
                            eState := eHold;
                        ELSE
                            bDoAdvance := TRUE;
                        END_IF
                    END_IF
                END_IF

            END_IF

        eHold:
            (* 单步推进：真正的换步在段 6 统一执行，此处只发请求 *)
            (* Advance request only, the actual switch happens in stage 6 *)
            IF fbTrigAdvance.Q THEN
                bDoAdvance := TRUE;
            END_IF

        eDone:
            (* 全部完成：启动沿可直接重新开始一轮 *)
            (* All done: a start edge begins a new cycle *)
            IF fbTrigStart.Q THEN
                nStep         := 0;
                bArmStep      := TRUE;
                bMaskNext     := TRUE;
                eState        := eRun;
            END_IF

        eFault:
            (* 故障锁存：保持步号便于现场定位，停用超时监控避免二次触发 *)
            (* Fault latched: the step index is kept for diagnosis, the timer is disarmed *)
            bTimeoutArmed := FALSE;

        ELSE
            (* 非法状态拦截：转故障并上报，不做隐式恢复 *)
            (* Illegal state interception: go to fault and report, no implicit recovery *)
            eState     := eFault;
            nFaultStep := nStep;
            uErrorId   := 16#0001_0005;

    END_CASE;

END_IF

(*------------------------------------------------------------------------------
 * 段 6｜推进执行（边界 B8）：末步完成进完成态并保持末步步号，其余步号加一
 *      Advance: the last step completes the sequence, otherwise the index increments
 *      推进只在此处发生一次，避免多处写步号造成跳步
 *      The index changes in exactly one place, which rules out double-stepping
 *-----------------------------------------------------------------------------*)
IF bDoAdvance THEN

    IF nStep >= (DL_SEQ_MAX_STEPS - 1) THEN
        eState := eDone;
    ELSE
        nStep      := nStep + 1;
        bMaskNext  := TRUE;
        bArmStep   := TRUE;
        eState     := eRun;
    END_IF

END_IF

(*------------------------------------------------------------------------------
 * 段 7｜步超时装载（边界 B3/B11）：进入新步时取该步超时并钳位
 *      Step timeout load: read and clamp the timeout when a step is entered
 *      超时为 0 表示该步不监控，挂死风险由调用方自担（手册明示）
 *      A zero timeout disables monitoring for that step, the caller carries the risk
 *-----------------------------------------------------------------------------*)
IF bArmStep THEN
    IF (nStep >= 0) AND (nStep < DL_SEQ_MAX_STEPS) THEN
        IF auStepTimeout[nStep] > DL_SEQ_TOUT_MAX THEN
            tEffTimeout   := DL_SEQ_TOUT_MAX;
            bTimeoutArmed := TRUE;
            uErrorId      := 16#0001_0001;
        ELSIF auStepTimeout[nStep] <= T#0S THEN
            tEffTimeout   := T#0S;
            bTimeoutArmed := FALSE;
        ELSE
            tEffTimeout   := auStepTimeout[nStep];
            bTimeoutArmed := TRUE;
        END_IF
    ELSE
        tEffTimeout   := T#0S;
        bTimeoutArmed := FALSE;
    END_IF
END_IF

(*------------------------------------------------------------------------------
 * 段 8｜输出刷新（边界 B8）：步号与状态标志集中在此一次赋值
 *      Output refresh: the step index and the status flags are written once here
 *-----------------------------------------------------------------------------*)
nCurrentStep := nStep;
bRunning     := (eState = eRun);
bDone        := (eState = eDone);
bError       := (eState = eFault);
tStepElapsed := fbTonStep.ET;

(*------------------------------------------------------------------------------
 * 段 9｜换步屏蔽标志提交（边界 B2）：本周期置的请求在下一周期生效并自动解除
 *      Mask commit: a request raised this scan takes effect next scan and self-clears
 *      这样换步后的第一个完整周期既不推进也不计时，旧步残留完成位无从生效
 *      The first full scan after a switch neither advances nor times, so stale bits die here
 *-----------------------------------------------------------------------------*)
bJustAdvanced := bMaskNext;
bMaskNext     := FALSE;
END_FUNCTION_BLOCK

(* ---- FB_DL_StepTimeRecorder.st ---- *)
(*==============================================================================
 * 组件名称 (Component)  : FB_DL_StepTimeRecorder
 * 所属子库 (Sublibrary) : DL_Base
 * 当前版本 (Version)    : 1.0.0
 * 兼容性 (Platform)     : CODESYS 3.5+ / TwinCAT 3 / 汇川 InoProShop / 施耐德 Machine Expert
 *                         仅依赖 Standard.library（R_TRIG），零厂商私有库
 * 功能描述 (Function)   : 顺控各步耗时在线采集统计（测量侧）。调用方每拍给出
 *                         当前激活步号 nStepId（0 = 无激活步），本件按扫描周期
 *                         tScan 对激活步做时间积分：步切换沿（步号变化或回 0）
 *                         时把累计时长入档（步号槽位记录 count/sum/last/min/max，
 *                         并派生 avg）。批量产线节拍分析、顺控瓶颈定位场景。
 * 来源标签 (Origin)     : 自研线（IEC 61131-3 标准语义的道莅防御性实现，clean-room）
 * 分工声明 (Pairing)    : StepTimeRecorder（测量侧，本件）↔ FB_DL_StepSequencer
 *                         （编排侧，既有件）：本件只消费步号快照做耗时统计，
 *                         不产生步进命令、不干预顺控相位、不持有步状态机
 *                         （R298 属主边界：测量不改编排）。
 * 边界语义 (Boundary)   : ① 步号闸：nStepId 落于 1..16 域外按 0（无激活步）处理
 *                         并置信息级 nWarnCnt 递增（越界钳位，R308 口径）；
 *                         ② 档位满：单步 count 达 DINT 上限饱和不再递增（防回绕，
 *                         上限 2^30 远超工程寿命，sum 同步饱和）；
 *                         ③ 除零防御：avg 仅在 count >= 1 时派生，除子恒 >= 1；
 *                         ④ 组态闸：tScan <= T#0S → bError 锁存（积分失真）；
 *                         ⑤ 监视型无主状态机（R23 周期监视型公约），无 CASE 相。
 * 来源标签 (Origin)     : T0 语义件；本件为自研线补口件，无 T0 对应条目。
 * 码位     (Codes)      : 按 R297 范式零 16# 码位硬编码；错误出口 BOOL(bError)，
 *                         码位待主控收口统一派号。
 * 红线自检 (Redline)    : 7 项红线已自检：R1 零全局 ✓｜R2 零物理地址 ✓｜R3 纯 IEC ✓
 *                         R4 越界钳位/饱和防回绕/除零防御 ✓｜R5 双语同行注释 ✓
 *                         R6 N/A（监视型无状态机，判据纯派生）✓
 *                         R7 R_TRIG 段 0 无条件每拍刷新 ✓
 * 验收向量 (Acceptance) : V1 步 3 激活 2.0s 后切步 → aStepLast[3]=2.0，
 *                         aStepAvg[3]=2.0，aStepCnt[3]=1；
 *                         V2 步 3 再测 3.0s → aStepAvg[3]=2.5，aStepMax[3]=3.0；
 *                         V3 nStepId=99 → 按 0 处理且 nWarnCnt 递增；
 *                         V4 bReset 上升沿全档清零（上电回夹防线）。
 * 修订历史 (Revision)   : 2026-11-20  v1.0.0  R49 首版（批 1 · 序号 5）
 *==============================================================================*)
FUNCTION_BLOCK FB_DL_StepTimeRecorder
VAR_INPUT
    nStepId  : INT := 0;                     (* 当前激活步号，0 = 无激活步，域 1..16 域外按 0 [步] / Active step id, 0 = none *)
    tScan    : TIME := T#10MS;               (* 扫描周期（积分步长），域 > T#0S [ms] / Scan cycle integration step *)
    bEnable  : BOOL := TRUE;                 (* 采集使能，FALSE 时冻结不积分不切档 [-] / Enable, FALSE freezes accumulation *)
    bReset   : BOOL := FALSE;                (* 复位命令，上升沿清全部档位与告警计数 [-] / Reset, rising edge clears all banks *)
END_VAR
VAR_OUTPUT
    aStepCnt  : ARRAY[1..16] OF DINT;        (* 各步样本计数（档位量）[个] / Sample count per step bank *)
    aStepLast : ARRAY[1..16] OF LREAL;       (* 各步最近一次耗时 [s] / Last duration per step *)
    aStepAvg  : ARRAY[1..16] OF LREAL;       (* 各步平均耗时 = sum/count [s] / Average duration per step *)
    aStepMin  : ARRAY[1..16] OF LREAL;       (* 各步最小耗时 [s] / Minimum duration per step *)
    aStepMax  : ARRAY[1..16] OF LREAL;       (* 各步最大耗时 [s] / Maximum duration per step *)
    bBanked   : BOOL;                        (* 本拍完成一次入档的单拍脉冲 [-] / Single-scan bank-update pulse *)
    nBankedId : INT;                         (* 最近入档步号（诊断镜像）[步] / Last banked step id *)
    nWarnCnt  : UDINT;                       (* 非法步号拒收累计（信息级台账）[次] / Illegal id rejection counter *)
    bError    : BOOL;                        (* 组态故障锁存标志（tScan 非法）[-] / Config fault latch flag *)
END_VAR
VAR
    rtReset  : R_TRIG;                       (* 复位沿实例，段 0 无条件调用 / Reset edge instance *)
    i        : INT;                          (* 复位清档循环游标 [-] / Reset clear loop cursor *)
    _nPrevId : INT;                          (* 上拍激活步号（切换沿检测基准）[步] / Previous active step id *)
    _fAccS   : LREAL;                        (* 当前步累计时长（积分器）[s] / Current step accumulator *)
    _fScanS  : LREAL := 0.01;                (* 扫描周期秒值缓存（TIME 秒换算）[s] / Scan cycle seconds cache *)
    _nCurId  : INT;                          (* 防御后生效步号（钳位结果）[步] / Sanitized current step id *)
    _bFault  : BOOL;                         (* 组态故障锁存位 / Config fault latch bit *)
END_VAR
VAR CONSTANT
    DL_ST_NMAX   : INT   := 16;              (* 步号容量上限（越界钳位目标）[步] / Step capacity limit *)
    DL_ST_DMAX   : DINT  := 1073741824;      (* 计数饱和上限 2^30（防回绕）[个] / Count saturation limit 2^30 *)
    DL_ST_SUMMAX : LREAL := 1.0E15;          (* 累计和饱和上限（防精度坍缩）[s] / Sum saturation limit *)
END_VAR

(* —— 段 0：当拍判据派生 + 沿实例无条件刷新（R228A） —— *)
rtReset(CLK := bReset);                                      (* 复位沿每拍必调 / Reset edge every scan *)
_fScanS := TIME_TO_LREAL(tScan) / 1000.0;                    (* 毫秒口径换算秒（舍入意图：整毫秒无损）[s] / Convert ms to seconds *)
IF _fScanS <= 1.0E-9 OR (tScan <= T#0S) THEN                 (* 组态闸：步长非法（含 TIME 下溢） / Config gate: illegal step *)
    _bFault := TRUE;                                         (* 锁存组态故障 / Latch config fault *)
END_IF

(* —— 段 1：单拍量预清零（锁存量与档位不入清单，R107） —— *)
bBanked := FALSE;                                            (* 入档单拍位预清，唯一分支置位 / Bank pulse preset *)

(* —— 段 2：复位沿处理（作用域：清故障 + 清全部档位数组 + 清积分器 + 清台账，R283 逐项声明） —— *)
IF rtReset.Q THEN
    _bFault := FALSE;                                        (* 清组态故障 / Clear config fault *)
    _fAccS := 0.0;                                           (* 清积分器 / Clear accumulator *)
    _nPrevId := 0;                                           (* 清上拍步号 / Clear previous id *)
    nWarnCnt := 0;                                           (* 清拒收台账 / Clear rejection counter *)
    nBankedId := 0;                                          (* 清入档镜像 / Clear banked mirror *)
    FOR i := 1 TO DL_ST_NMAX DO                              (* 全档位清零（上电回夹防线） / Clear all banks *)
        aStepCnt[i] := 0;                                    (* 清计数 / Clear count *)
        aStepLast[i] := 0.0;                                 (* 清最近值 / Clear last *)
        aStepAvg[i] := 0.0;                                  (* 清均值 / Clear avg *)
        aStepMin[i] := 0.0;                                  (* 清最小值 / Clear min *)
        aStepMax[i] := 0.0;                                  (* 清最大值 / Clear max *)
    END_FOR
END_IF

(* —— 段 3：步号钳位与非法拒收（域外按 0 处理，越界不越界访问，R308） —— *)
_nCurId := nStepId;                                          (* 生效步号初值 / Sanitized id init *)
IF (_nCurId < 1) OR (_nCurId > DL_ST_NMAX) THEN
    IF nStepId <> 0 THEN                                     (* 非零非法步号才记拒收（0 是合法空步） / Only nonzero illegal ids counted *)
        nWarnCnt := nWarnCnt + 1;                            (* 信息级台账递增（不置 bError，R90 信息级口径） / Info-level counter, not fault *)
    END_IF
    _nCurId := 0;                                            (* 按 0 处理 / Treat as none *)
END_IF

(* —— 段 4：激活积分 + 切换沿入档（监视型纯派生，无 CASE 相） —— *)
IF bEnable AND NOT _bFault THEN
    IF _nCurId = _nPrevId THEN
        IF _nCurId > 0 THEN
            _fAccS := _fAccS + _fScanS;                      (* 同步持续：积分累计（饱和防精度坍缩） / Same step: integrate *)
            IF _fAccS > DL_ST_SUMMAX THEN
                _fAccS := DL_ST_SUMMAX;                      (* 累计和饱和 / Saturate accumulator *)
            END_IF
        END_IF
    ELSE
        (* 切换沿：上一激活步收档（_nPrevId > 0 且累计 > 0 才入档，剔除断使能残片） / Step change: bank previous step *)
        IF (_nPrevId >= 1) AND (_nPrevId <= DL_ST_NMAX) AND (_fAccS > 0.0) THEN
            aStepLast[_nPrevId] := _fAccS;                   (* 记最近耗时 / Store last duration *)
            IF aStepCnt[_nPrevId] < DL_ST_DMAX THEN
                aStepAvg[_nPrevId] := (aStepAvg[_nPrevId] * DINT_TO_LREAL(aStepCnt[_nPrevId]) + _fAccS) / DINT_TO_LREAL(aStepCnt[_nPrevId] + 1);   (* 增量均值 = (旧和 + 新值)/(旧计数+1)，除子恒 >= 1 / Incremental mean, divisor >= 1 *)
                aStepCnt[_nPrevId] := aStepCnt[_nPrevId] + 1;   (* 计数递增（回绕防护） / Increment count, wrap-guarded *)
            END_IF
            IF (aStepMin[_nPrevId] <= 0.0) OR (_fAccS < aStepMin[_nPrevId]) THEN
                aStepMin[_nPrevId] := _fAccS;                (* 最小值更新（首样本或更小） / Min update *)
            END_IF
            IF _fAccS > aStepMax[_nPrevId] THEN
                aStepMax[_nPrevId] := _fAccS;                (* 最大值更新 / Max update *)
            END_IF
            bBanked := TRUE;                                 (* 入档单拍脉冲 / Bank pulse *)
            nBankedId := _nPrevId;                           (* 入档步号镜像 / Banked id mirror *)
        END_IF
        _fAccS := 0.0;                                       (* 新步积分器清零重开 / Reset accumulator for new step *)
        _nPrevId := _nCurId;                                 (* 更新切换基准 / Update change reference *)
    END_IF
END_IF

(* —— 段 5：出口映射（R191：bError 与 _bFault 名实同源） —— *)
bError := _bFault;                                           (* 组态故障镜像 / Config fault mirror *)
END_FUNCTION_BLOCK
